(* IEC 61131-3 sources: daoli-st-library/DL_Device (part 11) *)

(* ---- FC_DL_UpsLoadRateCalc.st ---- *)
(*
 * FC_DL_UpsLoadRateCalc | C1 | DL_Device
 * 功能：UPS 负载率、N+1 冗余下的最大允许负载率与过载判定       单位：功率 [kW]、负载率 [%]、台数 [台]
 * 工况边界：模块均分假设（各模块容量相同、均流良好）；额定功率须 >0、模块数须 ≥1、冗余台数须满足 0 ≤ nRedundant < nModules；不含电池放电与效率修正
 * 代数值回代：rated=400 kW、nModules=4、nRedundant=1 → maxPct=3/4×100=75 %、允许 300 kW；load=320 kW → 320>300 → xOverload=TRUE、负载率 80 %（与 spec 回代行一致）
 * 开源溯源：clean-room 自研，未复制任何第三方代码（无外部来源）
 *)
FUNCTION FC_DL_UpsLoadRateCalc : BOOL
VAR_INPUT
    rLoadKw     : REAL := 320.0;     // 实际负载功率 | actual load power [kW]
    rRatedKw    : REAL := 400.0;     // UPS 额定功率（全模块）| UPS rated power, all modules [kW]
    nModules    : INT := 4;          // 模块总数 | total module count [台]
    nRedundant  : INT := 1;          // 冗余模块数 | redundant module count [台]
END_VAR
VAR_OUTPUT
    rLoadRatePct     : REAL;         // 负载率 | load rate [%]
    rMaxPermittedPct : REAL;         // 冗余约束下的最大允许负载率 | maximum permitted load rate under the redundancy constraint [%]
    rMaxPermittedKw  : REAL;         // 冗余约束下的最大允许负载功率 | maximum permitted load power [kW]
    xOverload        : BOOL;         // 过载（超过冗余允许值）| overload beyond the redundancy allowance
    xRedundancyOk    : BOOL;         // 冗余成立（去冗余后仍有 ≥1 台可用）| redundancy valid, at least one module remains
    xValid           : BOOL;         // 输出有效 | outputs valid
END_VAR
VAR
    xFinLoad : BOOL;                 // 负载功率有限性 | load power is finite
    xFinRated: BOOL;                 // 额定功率有限性 | rated power is finite
    nUsable  : INT;                  // 允许带载的模块数（去冗余）| usable modules after removing the redundancy [台]
    rModules : REAL;                 // 模块数实数形式 | module count as a real number [台]
END_VAR
VAR CONSTANT
    DL_ULR_PCT : REAL := 100.0;      // 百分数换算系数 | percentage factor [%]
    DL_ULR_MIN : REAL := 1.0E-9;     // 额定功率下限（防零除）| rated power lower bound [kW]
END_VAR

// 段1｜非有限闸（R19）
xFinLoad := (rLoadKw = rLoadKw) AND ((rLoadKw - rLoadKw) = 0.0);
xFinRated := (rRatedKw = rRatedKw) AND ((rRatedKw - rRatedKw) = 0.0);
IF (NOT xFinLoad) OR (NOT xFinRated) THEN
    rLoadRatePct := 0.0;             // 安全值：负载率 0 | safe value, zero load rate
    rMaxPermittedPct := 0.0;
    rMaxPermittedKw := 0.0;
    xOverload := TRUE;               // 安全值：判过载，禁止新增负载 | safe value, flagged as overload
    xRedundancyOk := FALSE;
    xValid := FALSE;
    FC_DL_UpsLoadRateCalc := FALSE;
    RETURN;
END_IF

// 段2｜域闸：额定功率入分母须 >0，模块数与冗余数须自洽
IF (rRatedKw <= DL_ULR_MIN) OR (nModules < 1) OR (nRedundant < 0) OR (nRedundant >= nModules) THEN
    rLoadRatePct := 0.0;
    rMaxPermittedPct := 0.0;
    rMaxPermittedKw := 0.0;
    xOverload := TRUE;
    xRedundancyOk := FALSE;
    xValid := FALSE;
    FC_DL_UpsLoadRateCalc := FALSE;
    RETURN;
END_IF

// 段3｜算法：maxPct = (n−nRed)/n×100；负载率 = load/rated×100
nUsable := nModules - nRedundant;
rModules := INT_TO_REAL(nModules);
rMaxPermittedPct := INT_TO_REAL(nUsable) / rModules * DL_ULR_PCT;
rMaxPermittedKw := rRatedKw * INT_TO_REAL(nUsable) / rModules;
rLoadRatePct := rLoadKw / rRatedKw * DL_ULR_PCT;

// 段4｜判定：过载与冗余度（判据同源于原始功率与台数）
xOverload := rLoadKw > rMaxPermittedKw;
xRedundancyOk := nUsable >= 1;
xValid := TRUE;
FC_DL_UpsLoadRateCalc := TRUE;
END_FUNCTION

(* ---- FC_DL_VacHoldDecayChk.st ---- *)
(*
  ============================================================
  组件名 : FC_DL_VacHoldDecayChk
  分类   : DL_Device
  功能   : 真空保持衰减校验，按保持时段内的真空度跌落求衰减率并给出泄漏报警
  复杂度 : C1
  版本   : 1.0.0
  作者   : 道莅工业代码库工厂 / R81
  日期   : 2026-11-24
  开源溯源 : clean-room（no upstream）—— 依据公开工程公式自研，未复制任何上游实现
  红线自检 : R1 无GVL/R2 无物理地址/R3 纯IEC/R4 防除零/R5 双语注释
  接口说明 :
      衰减率 = (起始真空度 - 当前真空度) / 保持时长，单位 kPa/s。
      当前真空度高于起始值属测量异常或补抽工况，衰减率按 0 处理并置 bSuspect 提示，不判泄漏。
      衰减率严格大于允许限值才置泄漏报警，等于限值视为边界可控。
  ============================================================
*)
FUNCTION FC_DL_VacHoldDecayChk : BOOL
VAR_INPUT
    bEnable     : BOOL; // 使能：TRUE 时校验 / Enable: TRUE to check
    bErr        : BOOL; // 外部故障：TRUE 时立即退出并置结果无效 / External fault: TRUE aborts with invalid result
    rVacStart_kpa : REAL; // 保持时段起始真空度 [kPa] / vacuum level at the start of the hold phase [kilopascal]
    rVacNow_kpa : REAL; // 当前实测真空度 [kPa] / current measured vacuum level [kilopascal]
    rHoldTime_s : REAL; // 保持时段已持续时长 [s] / elapsed hold phase duration [second]
    rDecayLim   : REAL; // 允许的最大衰减率 [kPa/s] / permitted maximum decay rate [kilopascal per second]
END_VAR
VAR_OUTPUT
    rDecayRate : REAL; // 实测真空衰减率，负值按 0 处理 [kPa/s] / measured vacuum decay rate, negative clamped to zero [kilopascal per second]
    rDropKpa   : REAL; // 时段内真空度跌落量 [kPa] / vacuum drop within the hold phase [kilopascal]
    bLeakAlarm : BOOL; // 泄漏报警：TRUE 表示衰减率超过限值 / leak alarm, TRUE when the decay rate exceeds the limit
    bSuspect   : BOOL; // 数据可疑：TRUE 表示当前真空度高于起始值 / suspect data, TRUE when the current vacuum is above the start value
    bValid     : BOOL; // 输出有效：TRUE 表示结果可用 / Output valid
END_VAR
VAR CONSTANT
    DL_R_MAX   : REAL := 3.0E38;  // 实数上界，用于拦截 Inf [无量纲] / real upper bound used to reject infinity [dimensionless]
    DL_EPS     : REAL := 1.0E-12; // 除零判定阈值 [无量纲] / division guard threshold [dimensionless]
    DL_ZERO    : REAL := 0.0;     // 零值常量 [无量纲] / zero constant [dimensionless]
    DL_VAC_MAX : REAL := 101.3;   // 真空度物理上限，标准大气压 [kPa] / physical upper bound of the vacuum level, standard atmosphere [kilopascal]
END_VAR
VAR
    _bFin : BOOL := FALSE; // 输入有限性判定结果 / input finiteness verdict
END_VAR

    // 段 1｜出口预置：报警位保守置 FALSE，可疑位先置 FALSE
    rDecayRate := 0.0;
    rDropKpa := 0.0;
    bLeakAlarm := FALSE;
    bSuspect := FALSE;
    bValid := FALSE;
    // 段 2｜使能闸与外部故障闸
    IF NOT bEnable THEN
        RETURN;
    END_IF;
    IF bErr THEN
        RETURN;
    END_IF;
    // 段 3｜非有限闸
    _bFin := (rVacStart_kpa = rVacStart_kpa) AND (ABS(rVacStart_kpa) <= DL_R_MAX) AND (rVacNow_kpa = rVacNow_kpa) AND (ABS(rVacNow_kpa) <= DL_R_MAX) AND (rHoldTime_s = rHoldTime_s) AND (ABS(rHoldTime_s) <= DL_R_MAX) AND (rDecayLim = rDecayLim) AND (ABS(rDecayLim) <= DL_R_MAX);
    IF NOT _bFin THEN
        RETURN;
    END_IF;
    // 段 4｜域闸：保持时长严格为正，真空度与限值不得为负
    IF (ABS(rHoldTime_s) <= DL_EPS) OR (rHoldTime_s < DL_ZERO) THEN
        RETURN;
    END_IF;
    IF (rVacStart_kpa < DL_ZERO) OR (rVacNow_kpa < DL_ZERO) OR (rDecayLim < DL_ZERO) THEN
        RETURN;
    END_IF;
    IF (rVacStart_kpa > DL_VAC_MAX) OR (rVacNow_kpa > DL_VAC_MAX) THEN
        RETURN;
    END_IF;
    // 段 5｜跌落量与衰减率
    rDropKpa := rVacStart_kpa - rVacNow_kpa;
    IF rDropKpa < DL_ZERO THEN
        bSuspect := TRUE;
        rDropKpa := DL_ZERO;
        rDecayRate := DL_ZERO;
    ELSE
        bSuspect := FALSE;
        rDecayRate := rDropKpa / rHoldTime_s;
    END_IF;
    // 段 6｜泄漏报警
    IF rDecayRate > rDecayLim THEN
        bLeakAlarm := TRUE;
    ELSE
        bLeakAlarm := FALSE;
    END_IF;
    bValid := TRUE;
    FC_DL_VacHoldDecayChk := bValid;
END_FUNCTION

(* ---- FC_DL_VacuumGenDutyCalc.st ---- *)
(*
  ============================================================
  组件名 : FC_DL_VacuumGenDutyCalc
  分类   : DL_Device
  功能   : 真空发生器占空比计算，按单周期通电时长求占空比并折算压缩空气耗量
  复杂度 : C1
  版本   : 1.0.0
  作者   : 道莅工业代码库工厂 / R81
  日期   : 2026-11-24
  开源溯源 : clean-room（no upstream）—— 依据公开工程公式自研，未复制任何上游实现
  红线自检 : R1 无GVL/R2 无物理地址/R3 纯IEC/R4 防除零/R5 双语注释
  接口说明 :
      占空比 = 通电时长 / 循环周期 * 100，限幅 0~100。
      平均耗气量 = 额定耗气量 * 占空比 / 100，单位 L/min。
      通电时长超过循环周期属参数矛盾，判无效；周期为零则无法归一，同样判无效。
  ============================================================
*)
FUNCTION FC_DL_VacuumGenDutyCalc : BOOL
VAR_INPUT
    bEnable    : BOOL; // 使能：TRUE 时计算 / Enable: TRUE to compute
    bErr       : BOOL; // 外部故障：TRUE 时立即退出并置结果无效 / External fault: TRUE aborts with invalid result
    rOnTime_s  : REAL; // 单周期内真空发生器通电时长 [s] / generator energised time within one cycle [second]
    rCycle_s   : REAL; // 循环周期总时长 [s] / total cycle duration [second]
    rAirCons   : REAL; // 通电状态下的额定耗气量 [L/min] / rated air consumption while energised [litre per minute]
END_VAR
VAR_OUTPUT
    rDutyPct   : REAL; // 真空发生器占空比，限幅 0~100 [%] / generator duty cycle clamped to 0 to 100 [percent]
    rAirUseLpm : REAL; // 折算平均耗气量 [L/min] / equivalent average air consumption [litre per minute]
    bValid     : BOOL; // 输出有效：TRUE 表示结果可用 / Output valid
END_VAR
VAR CONSTANT
    DL_R_MAX   : REAL := 3.0E38;  // 实数上界，用于拦截 Inf [无量纲] / real upper bound used to reject infinity [dimensionless]
    DL_EPS     : REAL := 1.0E-12; // 除零判定阈值 [无量纲] / division guard threshold [dimensionless]
    DL_PCT     : REAL := 100.0;   // 百分数换算系数 [无量纲] / percentage scaling factor [dimensionless]
    DL_ZERO    : REAL := 0.0;     // 零值常量 [无量纲] / zero constant [dimensionless]
    DL_TOL_S   : REAL := 0.001;   // 时长比较容差 [s] / tolerance of the duration comparison [second]
    DL_CYC_MAX : REAL := 86400.0; // 循环周期合理上限，一天 [s] / sanity upper bound of the cycle duration, one day [second]
END_VAR
VAR
    _bFin : BOOL := FALSE; // 输入有限性判定结果 / input finiteness verdict
END_VAR

    // 段 1｜出口预置
    rDutyPct := 0.0;
    rAirUseLpm := 0.0;
    bValid := FALSE;
    // 段 2｜使能闸与外部故障闸
    IF NOT bEnable THEN
        RETURN;
    END_IF;
    IF bErr THEN
        RETURN;
    END_IF;
    // 段 3｜非有限闸
    _bFin := (rOnTime_s = rOnTime_s) AND (ABS(rOnTime_s) <= DL_R_MAX) AND (rCycle_s = rCycle_s) AND (ABS(rCycle_s) <= DL_R_MAX) AND (rAirCons = rAirCons) AND (ABS(rAirCons) <= DL_R_MAX);
    IF NOT _bFin THEN
        RETURN;
    END_IF;
    // 段 4｜域闸：周期严格为正且不超过一天，通电时长与耗气量非负
    IF (ABS(rCycle_s) <= DL_EPS) OR (rCycle_s < DL_ZERO) OR (rCycle_s > DL_CYC_MAX) THEN
        RETURN;
    END_IF;
    IF (rOnTime_s < DL_ZERO) OR (rAirCons < DL_ZERO) THEN
        RETURN;
    END_IF;
    // 段 5｜通电时长不得越过周期
    IF rOnTime_s > (rCycle_s + DL_TOL_S) THEN
        RETURN;
    END_IF;
    // 段 6｜占空比与限幅
    rDutyPct := rOnTime_s / rCycle_s * DL_PCT;
    IF rDutyPct < DL_ZERO THEN
        rDutyPct := DL_ZERO;
    END_IF;
    IF rDutyPct > DL_PCT THEN
        rDutyPct := DL_PCT;
    END_IF;
    // 段 7｜平均耗气量
    rAirUseLpm := rAirCons * rDutyPct / DL_PCT;
    bValid := TRUE;
    FC_DL_VacuumGenDutyCalc := bValid;
END_FUNCTION

(* ---- FC_DL_VacuumPadForceCalc.st ---- *)
(*
  ============================================================
  组件名 : FC_DL_VacuumPadForceCalc
  分类   : DL_Device
  功能   : 真空吸盘吸附力计算，由吸盘直径与真空度求理论吸附力并按安全系数折算可用力
  复杂度 : C1
  版本   : 1.0.0
  作者   : 道莅工业代码库工厂 / R81
  日期   : 2026-11-24
  开源溯源 : clean-room（no upstream）—— 依据公开工程公式自研，未复制任何上游实现
  红线自检 : R1 无GVL/R2 无物理地址/R3 纯IEC/R4 防除零/R5 双语注释
  接口说明 :
      吸附力 F = (pi/4) * (直径/1000)^2 * (真空度*1000)，直径先由 mm 折 m，真空度由 kPa 折 Pa，结果单位 N。
      可用力 = 理论力 / 安全系数；安全系数工程常用 1.5~3，低于 1.0 视为参数错误。
      面积同时以 mm2 输出，便于与样本册的吸盘规格直接对照。
  ============================================================
*)
FUNCTION FC_DL_VacuumPadForceCalc : BOOL
VAR_INPUT
    bEnable  : BOOL; // 使能：TRUE 时计算 / Enable: TRUE to compute
    bErr     : BOOL; // 外部故障：TRUE 时立即退出并置结果无效 / External fault: TRUE aborts with invalid result
    rDia_mm  : REAL; // 吸盘有效直径 [mm] / effective pad diameter [millimetre]
    rVacKpa  : REAL; // 工作真空度 [kPa] / working vacuum level [kilopascal]
    rSafety  : REAL; // 安全系数，常用 1.5~3 [无量纲] / safety factor, typically 1.5 to 3 [dimensionless]
END_VAR
VAR_OUTPUT
    rArea_mm2 : REAL; // 吸盘有效面积 [mm2] / effective pad area [square millimetre]
    rForceN   : REAL; // 理论吸附力 [N] / theoretical holding force [newton]
    rUsableN  : REAL; // 除以安全系数后的可用吸附力 [N] / usable holding force after the safety factor [newton]
    bValid    : BOOL; // 输出有效：TRUE 表示结果可用 / Output valid
END_VAR
VAR CONSTANT
    DL_PI      : REAL := 3.14159265; // 圆周率 [无量纲] / circular constant [dimensionless]
    DL_R_MAX   : REAL := 3.0E38;     // 实数上界，用于拦截 Inf [无量纲] / real upper bound used to reject infinity [dimensionless]
    DL_EPS     : REAL := 1.0E-12;    // 除零判定阈值 [无量纲] / division guard threshold [dimensionless]
    DL_MM_TO_M : REAL := 1000.0;     // 毫米折米系数 [mm/m] / millimetre to metre factor [millimetre per metre]
    DL_KPA_TO_PA : REAL := 1000.0;   // 千帕折帕系数 [Pa/kPa] / kilopascal to pascal factor [pascal per kilopascal]
    DL_QUARTER : REAL := 0.25;       // 四分之一，用于 pi/4 折算 [无量纲] / one quarter used for the pi over four term [dimensionless]
    DL_SAFE_MIN : REAL := 1.0;       // 安全系数下界 [无量纲] / lower bound of the safety factor [dimensionless]
    DL_SAFE_MAX : REAL := 10.0;      // 安全系数上界 [无量纲] / upper bound of the safety factor [dimensionless]
    DL_VAC_MAX : REAL := 101.3;      // 真空度物理上限，标准大气压 [kPa] / physical upper bound of the vacuum level, standard atmosphere [kilopascal]
END_VAR
VAR
    _bFin  : BOOL := FALSE; // 输入有限性判定结果 / input finiteness verdict
    _rDia  : REAL := 0.0;   // 吸盘直径折算米 [m] / pad diameter in metre [metre]
    _rArea : REAL := 0.0;   // 吸盘有效面积 [m2] / effective pad area [square metre]
    _rPress : REAL := 0.0;  // 压差折算帕 [Pa] / differential pressure in pascal [pascal]
END_VAR

    // 段 1｜出口预置
    rArea_mm2 := 0.0;
    rForceN := 0.0;
    rUsableN := 0.0;
    bValid := FALSE;
    // 段 2｜使能闸与外部故障闸
    IF NOT bEnable THEN
        RETURN;
    END_IF;
    IF bErr THEN
        RETURN;
    END_IF;
    // 段 3｜非有限闸
    _bFin := (rDia_mm = rDia_mm) AND (ABS(rDia_mm) <= DL_R_MAX) AND (rVacKpa = rVacKpa) AND (ABS(rVacKpa) <= DL_R_MAX) AND (rSafety = rSafety) AND (ABS(rSafety) <= DL_R_MAX);
    IF NOT _bFin THEN
        RETURN;
    END_IF;
    // 段 4｜域闸：直径严格为正且不超过 1 m，真空度为正且不超过大气压，安全系数在合理区间
    IF (ABS(rDia_mm) <= DL_EPS) OR (rDia_mm < 0.0) OR (rDia_mm > DL_MM_TO_M) THEN
        RETURN;
    END_IF;
    IF (ABS(rVacKpa) <= DL_EPS) OR (rVacKpa < 0.0) OR (rVacKpa > DL_VAC_MAX) THEN
        RETURN;
    END_IF;
    IF (rSafety < DL_SAFE_MIN) OR (rSafety > DL_SAFE_MAX) THEN
        RETURN;
    END_IF;
    // 段 5｜面积换算
    _rDia := rDia_mm / DL_MM_TO_M;
    _rArea := DL_PI * DL_QUARTER * _rDia * _rDia;
    rArea_mm2 := DL_PI * (rDia_mm * 0.5) * (rDia_mm * 0.5);
    // 段 6｜理论吸附力：面积乘压差
    _rPress := rVacKpa * DL_KPA_TO_PA;
    rForceN := _rArea * _rPress;
    // 段 7｜安全系数除前闸后再算可用力
    IF ABS(rSafety) <= DL_EPS THEN
        RETURN;
    END_IF;
    rUsableN := rForceN / rSafety;
    bValid := TRUE;
    FC_DL_VacuumPadForceCalc := bValid;
END_FUNCTION

(* ---- FC_DL_WinderTraversePitchCalc.st ---- *)
// FC_DL_WinderTraversePitchCalc v1.0.0
// 开源溯源：clean-room 自研（族 DL_Device，ST 生态实测 0 命中，无外部代码引入）
(*
  功能: 排线节距 = 带宽·(1 − 搭接率) [mm]；换向次数 = (卷绕线速·1000/60)/(2·排线行程) [次/min]；
        排线速度 = 节距·换向次数/60 [mm/s]。此为等比近似工程式：以排线行程近似替代卷径，
        适用于定行程往复排线的稳态估算，卷径变化需上层按卷径比修正。
  邻件/码位: 与 FC_DL_FiberDiameterFromDrawRateCalc 同属拉丝后端件（卷绕面 vs 直径面）；
             16#0002_9224 = 非有限、搭接率越界或带宽/行程/线速非正拒收。
*)
FUNCTION FC_DL_WinderTraversePitchCalc : REAL
VAR_INPUT
    fStrandWidth  : REAL := 20.0;   // 丝束带宽 [mm]，域 > 0 / Strand band width [mm]
    fOverlapRatio : REAL := 0.2;    // 搭接率 [-]，域 [0, 1) / Overlap ratio
    fWinderSpeed  : REAL := 900.0;  // 卷绕线速 [m/min]，域 > 0 / Winding speed [m/min]
    fTraverseLen  : REAL := 250.0;  // 排线行程 [mm]，域 > 0 / Traverse stroke [mm]
END_VAR
VAR_OUTPUT
    fPitch          : REAL;         // 排线节距 [mm] / Traverse pitch [mm]
    fTraverseSpeed  : REAL;         // 排线速度 [mm/s] / Traverse speed [mm/s]
    fReversalPerMin : REAL;         // 每分钟换向次数 [次/min] / Reversals per minute
    bValid          : BOOL;         // 结果有效回执 [-] / Result validity receipt
    uErrorId        : UDINT;        // 事件码，0 = 无事件 / Event code
END_VAR
VAR
    fSpeedMmS    : REAL := 0.0;     // 卷绕线速 [mm/s] / Winding speed [mm/s]
    fRoundTripMm : REAL := 0.0;     // 往返行程长度 [mm] / Round-trip travel [mm]
END_VAR
// 段 0：全路径出口安全缺省 / Safe defaults on all outlets
fPitch := 0.0;                      // 节距缺省零 / Pitch default zero
fTraverseSpeed := 0.0;              // 排线速度缺省零 / Traverse speed default zero
fReversalPerMin := 0.0;             // 换向次数缺省零 / Reversal rate default zero
bValid := FALSE;                    // 有效回执预清 / Validity preset clear
uErrorId := 16#0000;                // 事件码预清 / Event code preset clear
FC_DL_WinderTraversePitchCalc := 0.0;   // 返回值缺省零（镜像节距）/ Return default zero
// 段 1：非有限闸（四入参全枚举）/ Non-finite gate over all inputs
IF (fStrandWidth <> fStrandWidth) OR (fOverlapRatio <> fOverlapRatio)
   OR (fWinderSpeed <> fWinderSpeed) OR (fTraverseLen <> fTraverseLen)
   OR (ABS(fStrandWidth) >= 3.0E38) OR (ABS(fOverlapRatio) >= 3.0E38)
   OR (ABS(fWinderSpeed) >= 3.0E38) OR (ABS(fTraverseLen) >= 3.0E38) THEN
    uErrorId := 16#0002_9224;   // 入参非有限拒收 / Non-finite input reject
    RETURN;
END_IF
// 段 2：域闸（搭接率 [0,1) 防节距非正 + 带宽/行程/线速为正，R4）/ Domain gate
IF (fOverlapRatio < 0.0) OR (fOverlapRatio >= 1.0) THEN
    uErrorId := 16#0002_9224;   // 搭接率越界，节距将非正 / Overlap ratio out of range
    RETURN;
END_IF
IF (fStrandWidth <= 1.0E-6) OR (fTraverseLen <= 1.0E-6) OR (fWinderSpeed <= 1.0E-6) THEN
    uErrorId := 16#0002_9224;   // 带宽、行程或线速非正 / Non-positive width, stroke or speed
    RETURN;
END_IF
// 段 3：主计算（节距 → 换向次数 → 排线速度）/ Main computation
fPitch := fStrandWidth * (1.0 - fOverlapRatio);                 // 节距 [mm] / Pitch
fRoundTripMm := 2.0 * fTraverseLen;                             // 往返行程 [mm] / Round-trip travel
fSpeedMmS := fWinderSpeed * 1000.0 / 60.0;                      // 卷绕线速 [mm/s] / Winding speed
fReversalPerMin := fSpeedMmS / fRoundTripMm * 60.0;             // 换向次数 [次/min] / Reversal rate
fTraverseSpeed := fPitch * fReversalPerMin / 60.0;              // 排线速度 [mm/s] / Traverse speed
// 段 4：出口闸（三输出非有限复核 + 正数复核）/ Outlet gate
IF (fPitch <> fPitch) OR (fTraverseSpeed <> fTraverseSpeed) OR (fReversalPerMin <> fReversalPerMin)
   OR (ABS(fPitch) >= 3.0E38) OR (ABS(fTraverseSpeed) >= 3.0E38) OR (ABS(fReversalPerMin) >= 3.0E38)
   OR (fPitch <= 0.0) OR (fTraverseSpeed <= 0.0) THEN
    fPitch := 0.0;              // 复核失败回缺省 / Fallback on recheck failure
    fTraverseSpeed := 0.0;      // 复核失败回缺省 / Fallback on recheck failure
    fReversalPerMin := 0.0;     // 复核失败回缺省 / Fallback on recheck failure
    uErrorId := 16#0002_9224;   // 出口复核拒收 / Output recheck reject
    RETURN;
END_IF
bValid := TRUE;                 // 有效回执 / Validity receipt
FC_DL_WinderTraversePitchCalc := fPitch;    // 返回值镜像节距 / Return mirrors pitch
END_FUNCTION

(* ---- FB_DL_AdcNoiseFloorWatch.st ---- *)
(*
  ==================================================================
  组件名 Component  : FB_DL_AdcNoiseFloorWatch
  分类   Category   : DL_Device
  前缀   Naming     : FB_DL_ ｜ b/n/u/f/t/e/st 类型前缀制（R265）
  码位   Code ID    : 16#0003_071D / 071E（故障级）｜ 16#0003_071F / 0720（信息级）
  版本   Version    : 1.0.0
  复杂度 Complexity  : 中
  功能   Purpose    : ADC 测点底噪监视：静态期窗内标准差与上限比较（接地 / 屏蔽
                      劣化、前端供电噪声的早期征兆）。
  开源溯源 Origin    : 公开公式 clean-room，参考公开测量工程口径的底噪标准差判据
                      （分类与公式借鉴，零代码复制），本件实现、闸门与码位 100% 自有。
  许可证 License    : MIT
  参考   Reference  : IEC 61131-3:2013 §6.6 算术运算符；样本标准差（n−1 分母）
                      公开统计定义
  平台   Platform   : 纯 IEC 61131-3（FOR / 四则 / SQRT / TON 无），三平台通用
  依赖   Depends    : 仅 Standard.library（SQRT 属标准内建）
  分工声明 Split     : FB_DL_SignalFrozenDetect / FB_DL_SignalStuckWatch 监视
                      不变性；FB_DL_SignalStatistics 为通用统计出口；本件为静态期
                      噪声幅度监视（动静时序由 bStatic 外部给定），四件互引（R216）。
                      SQRT 原语经派单规格授权（窗内标准差属主口径）；统计内核委托
                      不适用（流式窗口件非整段数组口径，环窗驻留数据自算）。
  归属 Ownership     : 本件无 TYPE 声明；全部引脚为 IEC 标准原生类型。
  ------------------------------------------------------------------
  边界 Boundary     :
                      一 环形窗固定容量 256（禁动态分配）；活样本恒为下标
                         0.._nFill−1（写头仅在达 _nUse 时回卷，序不变量证明同族件）；
                         标准差与均值均为序不变量，回卷不影响结果；
                      二 bStatic 变更沿全窗清零（防静 / 动混合窗污染标准差口径）；
                         nWinLen 变更沿同样清窗；
                      三 标准差两遍法（均值先行、离差平方累加在后），禁「平方和减
                         均值平方」单遍式（灾难性抵消会产生负方差或 0，SPC 经典
                         事故，写死）；除子 DINT_TO_LREAL(_nFill − 1)：_nFill < 2 →
                         不计算（判据挂起，bValid = FALSE，除零防护，R61-D4 固化）；
                      四 fNoiseLim ≤ 0 或非有限 → 组态码 071D + 三件套 + RETURN
                         结构早退（族② 判据固化，R1 教训出厂即正确）；
                      五 fMeas 非有限 → 丢弃不入窗，nNonFinite 局部计数（不外显，
                         R62-D7 口径）超窗长一半 → 故障 071E + bValid = FALSE；
                      六 判据迟滞：fNoiseStd > fNoiseLim 触发，回落
                         < fNoiseLim×(1−fHystPct/100) 复原（两方向分别定义，R146）；
                      七 bEnable = FALSE 的语义写死（FB33-4 声明行）：判据复位 +
                         fNoiseStd 冻结（纯监视件，保留读数供 HMI）；
                      八 首拍 _bInit 全量初始化；无状态机（CASE N/A，R6 标注）；
                         无定时器 / 无边沿实例（段 0 无刷新对象）；无全局、无外部
                         变量、无物理地址。
  错误码 Codes      :
    16#0003_071D【故障级】组态非法（fNoiseLim ≤ 0 / 非有限；fHystPct < 0 / 非有限）
    16#0003_071E【故障级】测量失效（非有限样本累计超过窗长一半）
    16#0003_071F【信息级】底噪超上限（bNoiseHigh = TRUE）
    16#0003_0720【信息级】窗长越域已钳位（合法 16..256）
  码位反证 Note     :
    071D 与 071E 不可合并：071D 组态即刻判（与窗内容无关），071E 需窗已建立且坏点
    累计超半窗，处置人不同（组态工程师 / 仪表工），可由 nFill 与窗状态还原（R90）；
    071F / 0720 信息级与故障级分属不同子带（R75 子带纪律），不可跨用。
  验收 Acceptance   :
    算法已证（脚本）：未跑 ｜ 编译器已证（三平台）：未跑
    V1 恒定值 → std = 0、bNoiseHigh = FALSE
    V2 注入 ±0.5 方波抖动 → std ≈ 0.5，超限触发
    V3 限值上下 5% 波动（迟滞 10%）→ 不反复跳
    V4 fNoiseLim = 0 → 组态早退；V5 _nFill = 1 → 判据挂起 bValid = FALSE
    V6 bStatic 翻转 → 清窗 nFill = 0；V7 全 NaN → 故障 071E
  修订记录 Revision  :
    2026-11-21  v1.0.0  R63 首版（批 3 · 序号 9）
  ==================================================================
*)
FUNCTION_BLOCK FB_DL_AdcNoiseFloorWatch
VAR_INPUT
    bEnable   : BOOL := TRUE;  // 使能，FALSE 时判据复位 + 标准差冻结（边界七）/ the enable, false resets the criterion and freezes the std
    fMeas     : LREAL := 0.0;  // 测点实测值 [工程单位]，必须有限 / the measured value, must be finite
    bStatic   : BOOL := FALSE; // 静态期标志（过程稳态且无操作，由调用方给）[-] / the static period flag given by the caller
    nWinLen   : DINT := 64;    // 窗长 [个]，合法域 16..256，变更沿清窗 / the window length, legal sixteen to two hundred fifty six
    fNoiseLim : LREAL := 1.0;  // 底噪上限 [工程单位]，须 > 0 / the noise ceiling, must be positive
    fHystPct  : LREAL := 10.0; // 判据迟滞 [%]，须 ≥ 0 / the criterion hysteresis in percent, non negative
END_VAR
VAR_OUTPUT
    fNoiseStd  : LREAL := 0.0;           // 窗内标准差 [工程单位] / the window standard deviation
    bNoiseHigh : BOOL := FALSE;          // 底噪超限判据（带迟滞）[-] / the noise high criterion with hysteresis
    nFill      : DINT := 0;              // 窗填充数 [个] / the filled count
    bValid     : BOOL := FALSE;          // 判据可用 [-] / the criterion is usable
    eErr       : UDINT := 16#0000_0000;  // 错误码，0 = 正常 / the error code, zero is ok
    bError     : BOOL := FALSE;          // 故障标志（故障级码同拍置位，R45 配对）/ the fault flag raised with a fault level code
END_VAR
VAR
    _bInit     : BOOL := FALSE;              // 首拍初始化标志（R310 / FB50-2）/ the first scan flag
    _afWin     : ARRAY[0..255] OF LREAL;     // 采样环形窗 [工程单位]，固定容量 256 / the fixed capacity ring of samples
    _nHead     : DINT := 0;                  // 环形窗写头 [下标] / the ring write head
    _nFill     : DINT := 0;                  // 环形窗填充计数 [个] / the ring filled count
    _nUse      : DINT := 64;                 // 钳位后的窗长 [个] / the clamped window length
    _nUsePrev  : DINT := 0;                  // 上拍窗长快照 [个]，置 0 使首拍必触发清窗 / the previous length
    _bStaticPrev : BOOL := FALSE;            // 上拍静态期快照 [-] / the previous static flag
    _nClrIdx   : DINT := 0;                  // 清窗遍历索引 [下标] / the clearing traversal index
    _nSumIdx   : DINT := 0;                  // 统计遍历索引 [下标] / the statistics traversal index
    _nNonFinite: DINT := 0;                  // 非有限丢弃计数 [个]（仅局部留档，不外显，R62-D7 口径）/ the dropped non finite count, local only and never exposed
    _fSum      : LREAL := 0.0;               // 窗内样本和 [工程单位] / the window sample sum
    _fMean     : LREAL := 0.0;               // 窗内均值（两遍法第一遍）[工程单位] / the window mean of the first pass
    _fSqSum    : LREAL := 0.0;               // 离差平方和（两遍法第二遍）[工程单位²] / the squared deviation sum of the second pass
    _fStdUse   : LREAL := 0.0;               // 标准差工作副本 [工程单位] / the working standard deviation
    _fVar      : LREAL := 0.0;               // 样本方差（n−1 分母）[工程单位²] / the sample variance
    _bNoiseL   : BOOL := FALSE;              // 底噪超限迟滞状态（跨拍保持）/ the noise high hysteresis state
    _bCfgBad   : BOOL := FALSE;              // 组态非法标记（逐拍重算）/ the configuration fault flag
    _bWinClamp : BOOL := FALSE;              // 窗长钳位标记（逐拍重算，信息级 0720）/ the window clamp flag
    _bMeasBad  : BOOL := FALSE;              // 测量失效标记（逐拍重算）/ the measurement failure flag
    _bFinLim   : BOOL := FALSE;              // 上限有限闸结果（逐拍重算）/ the limit finiteness gate result
    _bFinHyst  : BOOL := FALSE;              // 迟滞有限闸结果（逐拍重算）/ the hysteresis finiteness gate result
    _bFinMeas  : BOOL := FALSE;              // 样本有限闸结果（逐拍重算）/ the sample finiteness gate result
END_VAR  // R64 结构补齐：VAR 段缺失的 END_VAR（门禁机械修复）
VAR CONSTANT
    DL_ANF_WMAX  : DINT := 256;      // 窗容量上界 [个]，与数组容量一致 / the capacity aligned with the array
    DL_ANF_WMIN  : DINT := 16;       // 窗长下界 [个] / the window floor
    DL_ANF_ZERO  : LREAL := 0.0;     // 实数零常量 [工程单位] / the real zero constant
    DL_ANF_PCT   : LREAL := 100.0;  // 百分比换算系数 [%] / the percentage scaling factor
    DL_ANF_ONE   : DINT := 1;        // 整型一常量 [个] / the integer one constant
    DL_ANF_TWO   : DINT := 2;        // 整型二常量 [个]（方差最少样本）/ the integer two constant, the minimum for a variance
    DL_ANF_ZEROI : DINT := 0;        // 整型零常量 [个] / the integer zero constant
    DL_ANF_HALF  : LREAL := 2.0;     // 半窗判据除子 [−] / the half window criterion divisor
END_VAR

// 段 0｜本件无定时器与边沿实例（纯统计监视器，R6 标注 N/A），无刷新对象 / segment 0, no timers and no edge instances exist here

// 段 1｜首拍初始化（FB50-2）/ segment 1, the first scan init
IF NOT _bInit THEN // 首拍一拍 / the first scan
    _bInit := TRUE; // 置首拍标志 / raise the first scan flag
    _nFill := DL_ANF_ZEROI; // 填充计数显式清零 / clear the filled count explicitly
    _nHead := DL_ANF_ZEROI; // 写头显式清零 / clear the write head explicitly
    _fSum := DL_ANF_ZERO; // 窗和显式清零 / clear the sum explicitly
    _nUsePrev := DL_ANF_ZEROI; // 窗长快照置 0，使段 3 变更沿必然触发一次清窗 / zero the snapshot so the change edge clears once
    _bStaticPrev := bStatic; // 静态期快照对齐首拍值（防首拍误清窗）/ align the static snapshot to avoid a spurious clear
    _bNoiseL := FALSE; // 迟滞状态显式清零 / clear the hysteresis state explicitly
    _nNonFinite := DL_ANF_ZEROI; // 非有限计数显式清零 / clear the non finite count explicitly
    FOR _nClrIdx := DL_ANF_ZEROI TO DL_ANF_WMAX - DL_ANF_ONE DO // 有界遍历全容量 / the bounded traversal over the full capacity
        _afWin[_nClrIdx] := DL_ANF_ZERO; // 窗元素逐项清零 / zero every window element
    END_FOR
END_IF

// 段 2｜组态域闸（边界四，族② 判据：全部限值逐个点名，R272）/ segment 2, the configuration gates
_bFinLim := (fNoiseLim = fNoiseLim) AND ((fNoiseLim - fNoiseLim) = (fNoiseLim - fNoiseLim)); // 上限有限 / the ceiling is finite
_bFinHyst := (fHystPct = fHystPct) AND ((fHystPct - fHystPct) = (fHystPct - fHystPct)); // 迟滞有限 / the hysteresis is finite
_bCfgBad := (NOT _bFinLim) OR (fNoiseLim <= DL_ANF_ZERO) OR (NOT _bFinHyst) OR (fHystPct < DL_ANF_ZERO); // 组态非法 / an illegal configuration
IF _bCfgBad THEN // 组态非法：结构早退（出口三件套 + RETURN，除法段不可达）/ an illegal configuration exits structurally
    fNoiseStd := _fStdUse; // 标准差取最近有效值 [工程单位]（禁自赋值出口，R261）/ the std takes the last valid value instead of a self assignment
    bNoiseHigh := FALSE; // 判据复位 / the criterion resets
    nFill := _nFill; // 填充计数照实出口 [个] / the fill count as is
    bValid := FALSE; // 判据不可用 / the criterion is not usable
    eErr := 16#0003_071D; // 故障级：组态非法 / fault grade, an illegal configuration
    bError := TRUE; // 同拍置故障标志（R45 配对）/ raise the fault flag on the same scan
    RETURN; // 结构早退 / the structural early exit
END_IF

// 段 3｜窗长钳位与变更沿 / 静态期变更沿全窗清零（边界二）/ segment 3, the window clamp and the change edge clears
_bWinClamp := FALSE; // 钳位标记预清零（单拍信息位，段 8 映射）/ preset the clamp flag false
_bMeasBad := FALSE; // 测量失效标记预清零 / preset the failure flag false
_nUse := nWinLen; // 窗长接管 [个] / take the window length
IF (_nUse < DL_ANF_WMIN) OR (_nUse > DL_ANF_WMAX) THEN // 窗长越域 / the length is out of the domain
    _bWinClamp := TRUE; // 置钳位标记（信息级 0720）/ raise the clamp flag
    IF _nUse < DL_ANF_WMIN THEN // 下界钳位 / the floor clamp
        _nUse := DL_ANF_WMIN; // 钳到下界 [个] / clamp to the floor
    ELSE // 上界钳位 / the ceiling clamp
        _nUse := DL_ANF_WMAX; // 钳到容量 [个] / clamp to the capacity
    END_IF
END_IF
IF (_nUse <> _nUsePrev) OR (bStatic <> _bStaticPrev) THEN // 窗长或静态期变更沿（含首拍）/ the length or the static flag changed
    _nHead := DL_ANF_ZEROI; // 写头回零 / reset the write head
    _nFill := DL_ANF_ZEROI; // 填充计数回零 / reset the filled count
    _fSum := DL_ANF_ZERO; // 窗和回零 / reset the sum
    _nNonFinite := DL_ANF_ZEROI; // 非有限计数回零 / reset the non finite count
    FOR _nClrIdx := DL_ANF_ZEROI TO DL_ANF_WMAX - DL_ANF_ONE DO // 有界遍历全容量 / the bounded traversal over the full capacity
        _afWin[_nClrIdx] := DL_ANF_ZERO; // 窗元素逐项清零（禁静动混合窗） / zero every element so no mixed window remains
    END_FOR
    _nUsePrev := _nUse; // 快照本拍窗长 / snapshot the length
    _bStaticPrev := bStatic; // 快照本拍静态期 / snapshot the static flag
END_IF

// 段 4｜失能分支：判据复位 + 标准差冻结（边界七声明行）/ segment 4, the disabled branch
IF NOT bEnable THEN // 失能 / disabled
    fNoiseStd := _fStdUse; // 标准差冻结最近有效值 [工程单位] / freeze the last valid std
    bNoiseHigh := FALSE; // 判据复位 / the criterion resets
    nFill := _nFill; // 填充计数照实出口 [个] / the fill count as is
    bValid := FALSE; // 失能即不可用 / the criterion is not usable while disabled
    bError := FALSE; // 失能不是故障 / a disabled device is not a fault
    eErr := 16#0000_0000; // 失能不发码 / no code is emitted while disabled
    RETURN; // 早退，窗保留 / early return with the window kept
END_IF

// 段 5｜样本入窗（非有限丢弃并计数，边界五）/ segment 5, push the sample or count the drop
_bFinMeas := (fMeas = fMeas) AND ((fMeas - fMeas) = (fMeas - fMeas)); // 样本有限 / the sample is finite
IF bStatic AND _bFinMeas THEN // 静态期且样本有限才入窗（动态期样本不进底噪窗）/ only a finite sample of a static period enters the noise window
    _fSum := _fSum - _afWin[_nHead] + fMeas; // 滑窗和更新 [工程单位] / update the sliding sum
    _afWin[_nHead] := fMeas; // 本拍样本入环 [工程单位] / push the sample
    _nHead := _nHead + DL_ANF_ONE; // 写头推进 / advance the head
    IF _nHead >= _nUse THEN // 回卷（按钳位窗长）/ wrap by the clamped length
        _nHead := DL_ANF_ZEROI; // 写头回零 / reset the head
    END_IF
    IF _nFill < _nUse THEN // 窗未满才累加 / count only while not full
        _nFill := _nFill + DL_ANF_ONE; // 填充计数推进 [个] / advance the filled count
    END_IF
ELSIF bStatic THEN // 静态期但样本非有限：丢弃计数 / a static period sample is broken, dropped and counted
    _nNonFinite := _nNonFinite + DL_ANF_ONE; // 非有限计数推进 [个] / advance the non finite count
END_IF
IF DINT_TO_LREAL(_nNonFinite) > (DINT_TO_LREAL(_nUse) / DL_ANF_HALF) THEN // 非有限累计超窗长一半（边界五）/ the non finite count exceeds half the window
    _bMeasBad := TRUE; // 置测量失效标记（码 071E）/ raise the failure flag
END_IF
nFill := _nFill; // 填充计数出口 [个] / the fill count outlet

// 段 6｜均值与标准差两遍法（边界三：除子 _nFill−1，_nFill < 2 判据挂起）/ segment 6, the two pass mean and standard deviation
IF _nFill >= DL_ANF_TWO THEN // 除子已证 ≥ 1（禁裸除子）/ the divisor is proven at least one
    _fMean := _fSum / DINT_TO_LREAL(_nFill); // 第一遍：窗均值 [工程单位] / the first pass mean
    _fSqSum := DL_ANF_ZERO; // 离差平方和清零 [工程单位²] / clear the squared deviation sum
    FOR _nSumIdx := DL_ANF_ZEROI TO _nFill - DL_ANF_ONE DO // 有界遍历活样本（上界已证 ≤ 256）/ the bounded traversal over the live samples
        _fSqSum := _fSqSum + ((_afWin[_nSumIdx] - _fMean) * (_afWin[_nSumIdx] - _fMean)); // 第二遍：离差平方累加 [工程单位²] / the second pass accumulates the squared deviations
    END_FOR
    _fVar := _fSqSum / DINT_TO_LREAL(_nFill - DL_ANF_ONE); // 样本方差（n−1 分母）[工程单位²] / the sample variance with the n minus one divisor
    IF _fVar < DL_ANF_ZERO THEN // 负方差兜底（两遍法下理论上不可达，防御保留）/ a negative variance, unreachable by theory, kept as a defence
        _fVar := DL_ANF_ZERO; // 方差钳零 [工程单位²] / clamp the variance to zero
    END_IF
    _fStdUse := SQRT(_fVar); // 标准差 [工程单位]，SQRT 属主口径见分工声明 / the standard deviation
ELSE // 样本不足：判据挂起 / too few samples, the criterion suspends
    fNoiseStd := _fStdUse; // 标准差保持最近有效值 [工程单位] / keep the last valid std
    bNoiseHigh := FALSE; // 判据复位 / the criterion resets
    bValid := FALSE; // 判据不可用（_nFill < 2，边界三）/ the criterion is not usable
    eErr := 16#0000_0000; // 挂起不是故障 / a suspension is not a fault
    bError := FALSE; // 无故障 / no fault
    RETURN; // 早退，禁除零 / early return, no division is reached
END_IF

// 段 7｜底噪判据迟滞（边界六，两方向分别定义，R146）/ segment 7, the noise criterion hysteresis
IF NOT _bNoiseL THEN // 未报警态 / the released state
    IF _fStdUse > fNoiseLim THEN // 超过上限 / above the ceiling
        _bNoiseL := TRUE; // 置迟滞状态 / set the hysteresis state
    END_IF
ELSE // 已报警态 / the tripped state
    IF _fStdUse < (fNoiseLim * (DL_ANF_PCT - fHystPct) / DL_ANF_PCT) THEN // 回落低于上限减迟滞 / below the ceiling minus the hysteresis
        _bNoiseL := FALSE; // 复原 / release
    END_IF
END_IF

// 段 8｜统一出口（单拍位映射 + 信息级重算，R187 / FB51-8）/ segment 8, the unified outlet
fNoiseStd := _fStdUse; // 标准差出口 [工程单位] / the std outlet
bNoiseHigh := _bNoiseL; // 判据出口（迟滞状态派生）/ the criterion outlet
bValid := (NOT _bMeasBad); // 判据可用（无测量失效）/ usable without a measurement failure
IF _bMeasBad THEN // 测量失效（故障级优先）/ the measurement failed
    bValid := FALSE; // 判据不可用 / the criterion is not usable
    bError := TRUE; // 故障位置位 / raise the fault bit
    eErr := 16#0003_071E; // 故障级：测量失效 / fault grade, the measurement failed
ELSIF _bNoiseL THEN // 底噪超限（信息级）/ the noise is high, informational
    bError := FALSE; // 信息级不置故障位 / the informational code never raises the fault bit
    eErr := 16#0003_071F; // 信息级：底噪超上限 / informational, the noise is over the ceiling
ELSIF _bWinClamp THEN // 窗长钳位（信息级）/ the length clamp, informational
    bError := FALSE; // 信息级不置故障位 / no fault bit
    eErr := 16#0003_0720; // 信息级：窗长越域已钳位 / informational, the length was clamped
ELSE // 无事件 / no event
    bError := FALSE; // 无故障 / no fault
    eErr := 16#0000_0000; // 正常 / ok
END_IF
END_FUNCTION_BLOCK

(* ---- FB_DL_AhuFilterDpBank.st ---- *)
// =====================================================================
// FB_DL_AhuFilterDpBank.st
// 空调箱 4 段过滤器压差四级分档（迟滞 + 各段独立去抖 + 低风量冻结）
// AHU 4-stage filter dP grading with per-stage debounce and hysteresis
// 所属子库: DL_Device    版本: v1.0.0    兼容: CODESYS V3.5+ / TwinCAT 3 / 汇川 InoProShop
// 码位: 16#0003_03D9 ~ 16#0003_03DD (本件独占 5 槽, 勿复用)
// 溯源: 道莅 clean-room 防御性实现
//       来源组标签: hvac, filter-monitoring, dp-grading, hysteresis, debounce
// 枚举属主: E_DL_FilterStage —— 本文件为全库唯一属主, 其他件只引用不重声明
// 修改记录: R30 初版 (ROUND_PLAN_R30 序 1, 由 R29 隔离底稿返修入册)
//           返修要点: 共享单实例去抖定时器改为 4 温区独立实例数组 aTonDeb,
//           每扫描周期无条件刷新全部 4 个 TON 实例, 候选作废显式复位;
//           任一区间切换去抖期间其他区间计时不被复位/冻结(验收点);
//           码位由作废段 03C5~03C9 重排为实测游标新段 03D9~03DD
// =====================================================================
// ---------------------------------------------------------------------
// 枚举定义: E_DL_FilterStage (全库唯一属主, 其他件只引用不重声明)
// ---------------------------------------------------------------------
TYPE E_DL_FilterStage :
(
    eClean,         // 洁净档 / Clean stage
    eEarly,         // 初堵档 / Early clog stage
    eMid,           // 中堵档 / Mid clog stage
    eChange,        // 更换档 / Change stage
    eSensorFault    // 传感器故障档 / Sensor fault stage
);
END_TYPE

FUNCTION_BLOCK FB_DL_AhuFilterDpBank
VAR_INPUT
    bEnable        : BOOL  := FALSE;   // 使能 / Enable
    afDp_Pa        : ARRAY[1..4] OF REAL;   // 各段压差 0~2000 Pa / Stage dP [Pa]
    afDpEarly_Pa   : ARRAY[1..4] OF REAL;   // 各段初堵阈值 10~500 Pa / Early clog threshold [Pa]
    afDpChange_Pa  : ARRAY[1..4] OF REAL;   // 各段更换阈值 20~1000 Pa / Change threshold [Pa]
    fHyst_Pa       : REAL  := 10.0;    // 迟滞回差 0~100 Pa / Hysteresis band [Pa]
    fDpMax_Pa      : REAL  := 1500.0;  // 传感器量程上限 >0 Pa / Sensor range limit [Pa]
    fFanPct        : REAL  := 0.0;     // 风机输出 0~100 百分比 / Fan duty [pct]
    fFanMinPct     : REAL  := 20.0;    // 判定最低风量 0~100 百分比 / Min fan duty for judging [pct]
    tDebounce      : TIME  := T#5S;    // 去抖时长 T#100MS~T#120S / Debounce duration [s]
END_VAR
VAR_OUTPUT
    aeStage        : ARRAY[1..4] OF E_DL_FilterStage;  // 各段档位 / Stage level per section
    auMaxStage     : USINT := 0;       // 全箱最高档 0~3 / Max stage of bank 0..3
    bChangeReq     : BOOL := FALSE;    // 更换请求 / Filter change required
    bFrozen        : BOOL := FALSE;    // 低风量冻结标志 / Frozen by low airflow
    eErr           : UDINT := 16#0003_03D9;  // 错误码 / Error code
END_VAR
VAR
    aTonDeb        : ARRAY[1..4] OF TON;   // 各段独立去抖定时器, 每拍无条件刷新 / Per-stage debounce timers, refreshed every cycle
    aPendStage     : ARRAY[1..4] OF E_DL_FilterStage;  // 各段候选档位 / Pending stage per section
    aPendActive    : ARRAY[1..4] OF BOOL;  // 各段候选有效标记 / Pending active flag per section
    eAbtCode       : UDINT := 16#0003_03D9;  // 本拍守卫闸中止码 / Abort code of this cycle
    bAbort         : BOOL := FALSE;    // 守卫闸中止标记 / Gate abort flag
    bSensorFlt     : BOOL := FALSE;    // 任一段传感器故障标记 / Any-stage sensor fault flag
    uZi            : INT   := 1;       // 1..4 数组下标 / Array subscript 1..4
    eTarget        : E_DL_FilterStage := E_DL_FilterStage.eClean;  // 本拍目标档 / Target stage this cycle
    uMaxTmp        : USINT := 0;       // 最高档临时量 / Max stage temporary
    tDebS          : REAL  := 0.0;     // 去抖秒值 / Debounce seconds [s]
    xFirstScan     : BOOL  := TRUE;    // 首扫标记 / First-scan flag
END_VAR

// ---------------------------------------------------------------------
// 代码位表（本件独占, 勿复用）:
//   16#0003_03D9 信息 分档正常
//   16#0003_03DA 故障 去抖时长非法或任一标量/数组输入非有限（本拍冻结保持, 非锁存, 恢复合法输入即解除）
//   16#0003_03DB 故障 阈值组态非法（量程上限不大于 0 或任一段初堵阈值不低于更换阈值）
//   16#0003_03DC 信息 低风量冻结（风机输出低于判定下限, 档位保持不推进）
//   16#0003_03DD 故障 任一段压差超量程或为负, 该段落传感器故障档
// ---------------------------------------------------------------------

// ---- 去抖秒值换算 / Debounce seconds conversion ----
tDebS := TIME_TO_REAL(tDebounce) / 1000.0;  // 毫秒换算秒 / Convert ms to seconds [s]

// ---- 守卫闸 1: 标量输入非有限与去抖时长合法域 / Gate 1: scalar finite and debounce range ----
bAbort    := FALSE;                 // 中止标记复位 / Reset abort flag
eAbtCode  := 16#0003_03D9;          // 中止码复位 / Reset abort code
IF (tDebounce = T#0MS) OR (tDebS < 0.1) OR (tDebS > 120.0)
   OR (fHyst_Pa <> fHyst_Pa) OR (ABS(fHyst_Pa) >= 1.0E12)
   OR (fDpMax_Pa <> fDpMax_Pa) OR (ABS(fDpMax_Pa) >= 1.0E12)
   OR (fFanPct <> fFanPct) OR (ABS(fFanPct) >= 1.0E12)
   OR (fFanMinPct <> fFanMinPct) OR (ABS(fFanMinPct) >= 1.0E12) THEN
    bAbort  := TRUE;                // 置中止 / Set abort
    eAbtCode := 16#0003_03DA;       // 码 03DA / Code 03DA
END_IF

// ---- 守卫闸 2: 逐段压差与阈值非有限判界 / Gate 2: per-stage finite check ----
IF NOT bAbort THEN
    FOR uZi := 1 TO 4 DO
        IF (afDp_Pa[uZi] <> afDp_Pa[uZi]) OR (ABS(afDp_Pa[uZi]) >= 1.0E12)
           OR (afDpEarly_Pa[uZi] <> afDpEarly_Pa[uZi]) OR (ABS(afDpEarly_Pa[uZi]) >= 1.0E12)
           OR (afDpChange_Pa[uZi] <> afDpChange_Pa[uZi]) OR (ABS(afDpChange_Pa[uZi]) >= 1.0E12) THEN
            bAbort   := TRUE;           // 置中止 / Set abort
            eAbtCode := 16#0003_03DA;   // 码 03DA / Code 03DA
        END_IF
    END_FOR
END_IF

// ---- 守卫闸 3: 阈值组态合法性 / Gate 3: threshold configuration ----
IF NOT bAbort THEN
    IF fDpMax_Pa <= 0.0 THEN
        bAbort   := TRUE;           // 量程非法 / Illegal range
        eAbtCode := 16#0003_03DB;   // 码 03DB / Code 03DB
    END_IF
END_IF
IF NOT bAbort THEN
    FOR uZi := 1 TO 4 DO
        IF afDpEarly_Pa[uZi] >= afDpChange_Pa[uZi] THEN
            bAbort   := TRUE;           // 阈值倒置 / Inverted thresholds
            eAbtCode := 16#0003_03DB;   // 码 03DB / Code 03DB
        END_IF
    END_FOR
END_IF

// ---- 首扫初始化 / First-scan initialization ----
IF xFirstScan THEN
    FOR uZi := 1 TO 4 DO
        aeStage[uZi]     := E_DL_FilterStage.eClean;    // 初始洁净档 / Init clean stage
        aPendStage[uZi]  := E_DL_FilterStage.eClean;    // 候选初始 / Pending init
        aPendActive[uZi] := FALSE;  // 候选无效 / Pending inactive
    END_FOR
    xFirstScan := FALSE;        // 清首扫标记 / Clear first-scan flag
END_IF

// ---- 低风量冻结与中止冻结推导 / Low-airflow freeze and abort freeze ----
IF bAbort THEN
    bFrozen := TRUE;            // 守卫闸中止按安全冻结处理 / Abort treated as safe freeze
ELSIF fFanPct < fFanMinPct THEN
    bFrozen := TRUE;            // 低风量冻结 / Low airflow freeze
ELSE
    bFrozen := FALSE;           // 正常非冻结 / Normal not frozen
END_IF

// ---- 逐段目标档计算与候选登记（不在此处调定时器）/ Per-stage target and pending registration ----
IF NOT bAbort AND NOT bFrozen THEN
    bSensorFlt := FALSE;        // 传感器故障标记复位 / Reset sensor fault flag
    bChangeReq := FALSE;        // 更换请求复位 / Reset change request
    FOR uZi := 1 TO 4 DO
        // 传感器故障判: 超量程或负压差 / Sensor fault: over-range or negative dP
        IF (afDp_Pa[uZi] > fDpMax_Pa) OR (afDp_Pa[uZi] < 0.0) THEN
            aeStage[uZi]     := E_DL_FilterStage.eSensorFault;  // 落传感器故障档 / Sensor fault stage
            aPendActive[uZi] := FALSE;  // 候选作废 / Pending void
            bSensorFlt := TRUE;         // 置传感器故障 / Set sensor fault
            bChangeReq := TRUE;         // 故障档也需现场处置 / Fault stage requests action
        ELSE
            // 双阈值迟滞分档: 严格大于阈值才切档, 恰好等于阈值保持原档 / Strict-greater hysteresis grading
            CASE aeStage[uZi] OF
                E_DL_FilterStage.eClean:        // 当前洁净 / Currently clean
                    IF afDp_Pa[uZi] > (afDpEarly_Pa[uZi] + fHyst_Pa) THEN
                        eTarget := E_DL_FilterStage.eEarly;     // 越升档阈值 → 初堵 / Above rise threshold
                    ELSE
                        eTarget := E_DL_FilterStage.eClean;     // 保持 / Hold
                    END_IF
                E_DL_FilterStage.eEarly:        // 当前初堵 / Currently early
                    IF afDp_Pa[uZi] > (afDpChange_Pa[uZi] + fHyst_Pa) THEN
                        eTarget := E_DL_FilterStage.eChange;    // 越更换阈值 / Above change threshold
                    ELSIF afDp_Pa[uZi] < (afDpEarly_Pa[uZi] - fHyst_Pa) THEN
                        eTarget := E_DL_FilterStage.eClean;     // 回落洁净 / Fall back clean
                    ELSE
                        eTarget := E_DL_FilterStage.eEarly;     // 保持 / Hold
                    END_IF
                E_DL_FilterStage.eMid:          // 当前中堵 / Currently mid
                    IF afDp_Pa[uZi] > (afDpChange_Pa[uZi] + fHyst_Pa) THEN
                        eTarget := E_DL_FilterStage.eChange;    // 越更换阈值 / Above change threshold
                    ELSIF afDp_Pa[uZi] < (afDpEarly_Pa[uZi] - fHyst_Pa) THEN
                        eTarget := E_DL_FilterStage.eClean;     // 回落洁净 / Fall back clean
                    ELSE
                        eTarget := E_DL_FilterStage.eMid;       // 保持 / Hold
                    END_IF
                E_DL_FilterStage.eChange:       // 当前更换档 / Currently change
                    IF afDp_Pa[uZi] < (afDpChange_Pa[uZi] - fHyst_Pa) THEN
                        eTarget := E_DL_FilterStage.eMid;       // 回落中堵 / Fall back mid
                    ELSE
                        eTarget := E_DL_FilterStage.eChange;    // 保持 / Hold
                    END_IF
                E_DL_FilterStage.eSensorFault:  // 故障档: 压差恢复量程内后按洁净档重新进入 / Fault holds, re-enter via grading
                    eTarget := E_DL_FilterStage.eClean;     // 目标回洁净档, 去抖后切换 / Target clean, switch after debounce
                ELSE                            // 非法档位拦截 / Illegal stage interception
                    eTarget := E_DL_FilterStage.eSensorFault;   // 落故障档 / Fall to fault stage
            END_CASE

            // 候选登记: 目标与当前不同才登记 / Register pending only if target differs
            IF eTarget <> aeStage[uZi] THEN
                IF (NOT aPendActive[uZi]) OR (aPendStage[uZi] <> eTarget) THEN
                    aPendStage[uZi]  := eTarget;    // 登记新候选 / Register new candidate
                    aPendActive[uZi] := TRUE;       // 候选有效 / Pending active
                END_IF
            ELSE
                aPendActive[uZi] := FALSE;      // 目标即当前档, 候选作废 / Target equals current, void
            END_IF
        END_IF

        // 更换档请求判 / Change stage request check
        IF aeStage[uZi] = E_DL_FilterStage.eChange THEN
            bChangeReq := TRUE;     // 任一段处于更换档 / Any stage at change
        END_IF
    END_FOR
ELSE
    bSensorFlt := FALSE;            // 冻结/中止拍不重推传感器判据 / No sensor re-judge on frozen cycle
    bChangeReq := FALSE;            // 冻结拍不置更换请求 / No change request on frozen cycle
END_IF

// ---- 4 个去抖定时器无条件周期刷新（本 FOR 循环每拍必执行全部 4 个实例,
//      不放进任何 IF 分支; 候选作废分支传 IN 为假显式复位而不是跳过调用）
//      Unconditional refresh of all 4 TON instances every cycle ----
FOR uZi := 1 TO 4 DO
    IF (NOT bAbort) AND (NOT bFrozen) AND aPendActive[uZi] AND (aPendStage[uZi] <> aeStage[uZi]) THEN
        aTonDeb[uZi](IN := TRUE, PT := tDebounce);  // 本拍继续计时 / Keep timing this cycle
        IF aTonDeb[uZi].Q THEN
            aeStage[uZi] := aPendStage[uZi];        // 去抖通过, 档位切换 / Switch after debounce
            aPendActive[uZi] := FALSE;              // 候选完成 / Pending done
        END_IF
    ELSE
        aPendActive[uZi] := FALSE;                  // 候选作废 / Pending void
        aTonDeb[uZi](IN := FALSE, PT := tDebounce); // 候选作废显式复位 / Explicit reset on void
    END_IF
END_FOR

// ---- 最高档统计（只统计非传感器故障段）/ Max stage excluding sensor-fault sections ----
uMaxTmp := 0;                   // 临时量复位 / Reset temporary
FOR uZi := 1 TO 4 DO
    IF aeStage[uZi] <> E_DL_FilterStage.eSensorFault THEN
        CASE aeStage[uZi] OF
            E_DL_FilterStage.eClean:    // 档 0 / Stage 0
                uMaxTmp := uMaxTmp;     // 保持 0 / Keep 0
            E_DL_FilterStage.eEarly:    // 档 1 / Stage 1
                IF uMaxTmp < 1 THEN
                    uMaxTmp := 1;       // 升到 1 / Raise to 1
                END_IF
            E_DL_FilterStage.eMid:      // 档 2 / Stage 2
                IF uMaxTmp < 2 THEN
                    uMaxTmp := 2;       // 升到 2 / Raise to 2
                END_IF
            E_DL_FilterStage.eChange:   // 档 3 / Stage 3
                uMaxTmp := 3;           // 升到 3 / Raise to 3
            ELSE                        // 兜底: 非法档不计入 / Fallback: illegal stage not counted
                uMaxTmp := uMaxTmp;     // 保持 / Keep
        END_CASE
    END_IF
END_FOR
auMaxStage := uMaxTmp;          // 输出最高档 / Output max stage

// ---- 错误码仲裁（每拍重算, 非锁存, 恢复合法输入即解除）/ Error arbitration recomputed each cycle ----
IF bAbort THEN
    eErr := eAbtCode;           // 守卫闸中止码优先 / Gate abort code first
ELSIF bSensorFlt THEN
    eErr := 16#0003_03DD;       // 传感器故障 / Sensor fault
ELSIF bFrozen THEN
    eErr := 16#0003_03DC;       // 低风量冻结 / Low airflow freeze
ELSE
    eErr := 16#0003_03D9;       // 分档正常 / Grading normal
END_IF

END_FUNCTION_BLOCK

(* ---- FB_DL_AirCompressorLoadUnload.st ---- *)
(*
  Name        : FB_DL_AirCompressorLoadUnload
  Category    : DL_Device
  Version     : 1.0.0
  Purpose     : 空压机加卸载调压：压力带双阈迟滞加卸载切换，加载最小驻留防短周期振荡，卸载超时置维护级告警不自动停机；/ Air compressor load/unload pressure control: dual-threshold hysteresis switching, minimum load dwell against short cycling, unload timeout raising a maintenance-level warning without auto stop
  溯源        : 借 lbp-basic-process 与行业池的调压组织，clean-room 实现
  Boundary    : ① 压力带组态闸：加载阈 < 卸载阈否则锁存故障（相等不立）；
                ② 双阈迟滞直比（加载阈/卸载阈比较，禁浮点等值）；
                ③ 卸载持续 > 卸载超时 → 置维护级告警（bMaintWarn 锁存至复位沿，不自动停机不迁故障相，属主边界）；
                ④ 加载最小驻留防短周期振荡：驻留期内卸载请求暂存不丢（驻留满即执行）；
                ⑤ 压力传感器非有限 → 保持当前负载态 + bSensorBad 当拍出口（不切态防误动作）；
                ⑥ 本件为命令层，不直接驱动接触器（属主边界，出加/卸载命令信号）。
*)
TYPE E_DL_AclState :
(
    eIdle   := 0,                            (* 未使能（命令全停） / Idle, commands off *)
    eLoad   := 10,                           (* 加载相 / Loading *)
    eUnload := 20,                           (* 卸载相 / Unloading *)
    eFault  := 90                            (* 故障锁存相 / Fault latched *)
);
END_TYPE

TYPE E_DL_AclCause :
(
    eNone      := 0,                         (* 无成因 / No cause *)
    eCfgIllegal:= 1,                        (* 组态非法：压力带阈值倒挂 / Illegal config *)
    eUnloadTime:= 2,                        (* 维护级：卸载超时（不置 bError，边界③） / Maintenance: unload timeout *)
    ePhaseBad  := 3                         (* 非法相位兜底 / Illegal phase fallback *)
);
END_TYPE

FUNCTION_BLOCK FB_DL_AirCompressorLoadUnload
VAR_INPUT
    fPress   : REAL := 0.0;                  (* 储气罐压力 [bar] / Receiver pressure *)
    fLoadTh  : REAL := 6.0;                  (* 加载阈（下限），域 < 卸载阈 [bar] / Load threshold *)
    fUnloadTh: REAL := 8.0;                  (* 卸载阈（上限）[bar] / Unload threshold *)
    tLoadMin : TIME := T#30S;                (* 加载最小驻留，域 > T#0S [ms] / Minimum load dwell *)
    tUnloadMax: TIME := T#10M;               (* 卸载超时，域 > T#0S [ms] / Unload timeout *)
    tScan    : TIME := T#100MS;              (* 扫描周期，域 > T#0S [ms] / Scan period *)
    bEnable  : BOOL := TRUE;                 (* 使能 [-] / Enable *)
    bReset   : BOOL := FALSE;                (* 复位命令，上升沿清故障与告警 [-] / Reset command *)
END_VAR
VAR_OUTPUT
    bLoadCmd : BOOL;                         (* 加载命令信号 [-] / Load command *)
    bUnloadCmd: BOOL;                        (* 卸载命令信号 [-] / Unload command *)
    bMaintWarn: BOOL;                        (* 维护级告警锁存（卸载超时，复位沿清，边界③）[-] / Maintenance warning latched *)
    bSensorBad: BOOL;                        (* 压力传感器失效当拍出口（边界⑤）[-] / Sensor bad outlet *)
    eState   : E_DL_AclState;                (* 状态出口 / State outlet *)
    eCause   : E_DL_AclCause;                (* 成因出口（R190 归因唯一） / Cause outlet *)
    bError   : BOOL;                         (* 故障锁存标志 [-] / Fault latch flag *)
END_VAR
VAR
    _eState : E_DL_AclState := E_DL_AclState.eIdle;  (* 内部相位（CASE 唯一写入目标） / Internal phase *)
    _eCause : E_DL_AclCause := E_DL_AclCause.eNone;  (* 成因锁存量 / Latched cause *)
    rtReset : R_TRIG;                        (* 复位沿实例，段 0 无条件调用 / Reset edge instance *)
    tonLoad : TON;                           (* 加载驻留计时（IN 串 eLoad 相闸，R40） / Load dwell timer *)
    tonUnl  : TON;                           (* 卸载持续计时（IN 串 eUnload 相闸，R40） / Unload duration timer *)
    _bFault : BOOL;                          (* 故障锁存位 / Latched fault bit *)
    _bCfgBad: BOOL;                          (* 组态非法当拍量 / Illegal config this scan *)
    _bFin   : BOOL;                          (* 压力有限性当拍量（边界⑤） / Pressure finiteness *)
    _bUnlReq: BOOL;                          (* 卸载请求暂存量（驻留期内不丢，边界④） / Buffered unload request *)
    _fDtSec : REAL;                          (* 扫描周期秒值（信息级备用派生）[s] / Scan period seconds *)
END_VAR
VAR CONSTANT
    DL_ACL_EPS : REAL := 1.0E-6;             (* 判零容差 [-] / Epsilon *)
END_VAR

(* —— 段 0：当拍判据派生 + 实例无条件刷新（R228A；TON 全段 0 无 IF 包裹，R40） —— *)
_bCfgBad := NOT (fLoadTh < fUnloadTh)                    (* 压力带组态闸：加载阈 < 卸载阈（边界①） / Band config gate *)
            OR (fLoadTh <= DL_ACL_EPS)                   (* 加载阈正域闸 / Load threshold gate *)
            OR NOT (tLoadMin > T#0S) OR NOT (tUnloadMax > T#0S) OR NOT (tScan > T#0S);   (* 周期域闸 / Period gates *)
rtReset(CLK := bReset);                                  (* 复位沿每拍必调 / Reset edge every scan *)
_bFin := (fPress = fPress) AND ((fPress - fPress) = (fPress - fPress));   (* 压力 NaN 自反 + Inf 差判闸（边界⑤） / Pressure NaN and Inf gate *)
_fDtSec := TIME_TO_LREAL(tScan) / 1000.0;                (* 扫描周期秒化（除子常量 1000） / Scan period seconds *)
tonLoad(IN := (_eState = E_DL_AclState.eLoad), PT := tLoadMin);          (* 加载驻留：相位闸 + 无条件调用（R40） / Load dwell timer *)
tonUnl(IN := (_eState = E_DL_AclState.eUnload), PT := tUnloadMax);       (* 卸载持续：相位闸 + 无条件调用（R40） / Unload timer *)

(* —— 段 1：单拍量预清零（R107） —— *)
bLoadCmd := FALSE;                                       (* 加载命令出口预清（派生拍覆盖） / Load command preset *)
bUnloadCmd := FALSE;                                     (* 卸载命令出口预清 / Unload command preset *)
bSensorBad := FALSE;                                     (* 传感器失效当拍出口预清 / Sensor bad preset *)

(* —— 段 2：复位沿处理（作用域：清故障 + 清维护告警 + 迁 eIdle，R283 逐项声明） —— *)
IF rtReset.Q THEN
    _bFault := FALSE;                                    (* 清故障锁存 / Clear fault *)
    _eCause := E_DL_AclCause.eNone;                      (* 清成因 / Clear cause *)
    bMaintWarn := FALSE;                                 (* 清维护告警锁存 / Clear maintenance warning *)
    _bUnlReq := FALSE;                                   (* 清卸载请求暂存 / Clear buffered request *)
    _eState := E_DL_AclState.eIdle;                      (* 迁未使能相 / Back to idle *)
END_IF

(* —— 段 3：组态故障锁存（锁存至复位沿，R189） —— *)
IF _bCfgBad AND NOT _bFault THEN
    _bFault := TRUE;                                     (* 锁存故障位 / Latch fault *)
    _eCause := E_DL_AclCause.eCfgIllegal;                (* 成因：组态非法 / Cause illegal config *)
    _eState := E_DL_AclState.eFault;                     (* 同步迁故障相 / Migrate to fault *)
END_IF

(* —— 段 4：CASE 主状态机（ELSE 兜底迁 eFault，红线 6） —— *)
CASE _eState OF
    E_DL_AclState.eIdle:                                 (* 未使能：命令全停确定值 / Idle *)
        bLoadCmd := FALSE;                               (* 失能加载命令 FALSE / Disabled load false *)
        bUnloadCmd := FALSE;                             (* 失能卸载命令 FALSE / Disabled unload false *)
        IF bEnable AND NOT _bFault THEN
            _eState := E_DL_AclState.eLoad;              (* 使能先入加载相（建压优先） / Enter loading *)
        END_IF
    E_DL_AclState.eLoad:                                 (* 加载相：驻留 + 双阈迟滞切换 / Loading *)
        IF NOT bEnable THEN
            _eState := E_DL_AclState.eIdle;              (* 失能回未使能 / Back to idle *)
        ELSIF NOT _bFin THEN
            bSensorBad := TRUE;                          (* 传感器失效：保持当前态（边界⑤） / Sensor bad hold *)
        ELSE
            IF fPress >= fUnloadTh THEN
                _bUnlReq := TRUE;                        (* 驻留期内卸载请求暂存不丢（边界④） / Buffer unload request *)
            END_IF
            IF tonLoad.Q AND _bUnlReq THEN               (* 驻留满 + 有暂存请求：迁卸载（边界④） / Dwell done and request *)
                _bUnlReq := FALSE;                       (* 请求消费清零 / Request consumed *)
                _eState := E_DL_AclState.eUnload;        (* 迁卸载相 / To unloading *)
            END_IF
        END_IF
    E_DL_AclState.eUnload:                               (* 卸载相：下阈回加载 + 超时维护告警 / Unloading *)
        IF NOT bEnable THEN
            _eState := E_DL_AclState.eIdle;              (* 失能回未使能 / Back to idle *)
        ELSIF NOT _bFin THEN
            bSensorBad := TRUE;                          (* 传感器失效：保持当前态（边界⑤） / Sensor bad hold *)
        ELSE
            IF tonUnl.Q THEN                             (* 卸载持续超时（边界③） / Unload timeout *)
                bMaintWarn := TRUE;                      (* 维护级告警锁存（复位沿清，不自动停机） / Maintenance warning latch *)
                _eCause := E_DL_AclCause.eUnloadTime;    (* 成因：卸载超时（信息级不置 bError，边界③） / Cause unload time *)
            END_IF
            IF fPress <= fLoadTh THEN                    (* 压力回落到加载阈：迁加载（双阈迟滞直比，边界②） / Back to load *)
                _eState := E_DL_AclState.eLoad;          (* 迁加载相 / To loading *)
            END_IF
        END_IF
    E_DL_AclState.eFault:                                (* 故障相：命令全停冻结，仅复位沿出 / Fault *)
        ;                                                (* 锁存回放（R28） / Replay from latch *)
    ELSE                                                 (* 非法相位兜底迁安全态 / Illegal phase fallback *)
        _eState := E_DL_AclState.eFault; _bFault := TRUE;    (* 迁故障相 + 同步锁存 / To fault and latch *)
        _eCause := E_DL_AclCause.ePhaseBad;              (* 成因：非法相位 / Cause illegal phase *)
END_CASE

(* —— 段 5：出口映射（名实双出口，R191；bError/eState 同源） —— *)
bLoadCmd := (_eState = E_DL_AclState.eLoad);             (* 加载命令 = 加载相镜像 / Load command mirror *)
bUnloadCmd := (_eState = E_DL_AclState.eUnload);         (* 卸载命令 = 卸载相镜像 / Unload command mirror *)
bError := _bFault;                                       (* 故障标志镜像 / Fault flag mirror *)
eState := _eState;                                       (* 状态出口 / State outlet *)
eCause := _eCause;                                       (* 成因出口 / Cause outlet *)
END_FUNCTION_BLOCK

(* ---- FB_DL_AirDryerDiag.st ---- *)
(*
  ==================================================================
  组件名 Component  : FB_DL_AirDryerDiag
  分类   Category   : DL_Device
  前缀   Naming     : FB_DL_ ｜ b/n/u/f/t/e/st 类型前缀制（R265）
  复杂度 Complexity  : 中
  版本   Version    : 1.0.0
  功能   Purpose    : 压缩空气干燥机诊断（露点越限 + 再生阀时序状态机 + 切换周期劣化档）。
  来源   Source     : t2-2-lbp（干燥机诊断公开工艺语义）
  平台   Platform   : 纯 IEC 61131-3（TON / R_TRIG / CASE / TIME_TO_DINT），三平台通用
  分工声明 Split     : 与 FB_DL_DryerProtect（停机保护属主，若在册）分工——本件
                      只做诊断与周期劣化分档，不做停机联锁（R216 双向互引）。
  作者   Author     : 道莅代码库 · PLC 编程专家（R61）
  归属 Ownership     : E_DL_DryerPhase 属主为本文件（全库唯一定义，R264）；
                      引用件只引用不重声明。
  ------------------------------------------------------------------
  边界 Boundary     :
                      一 露点非有限闸逐个点名（R272：fDewPnt / fDewLim /
                         fDeg1Ratio / fDeg2Ratio 四个浮点引脚逐个判）；
                      二 再生切换周期劣化分档阈值全提为输入（fDeg1Ratio /
                         fDeg2Ratio [-]，实测周期与名义周期之比阈值，R 红线 7）；
                         组态递增配比违反判组态锁存（070F）；
                      三 状态机 CASE 必带 ELSE 兜底（R25 批次教训）；TON /
                         R_TRIG 段 0 无条件刷新（禁入分支，R7）；
                      四 故障锁存解除式逐条自证：bReset 上升沿清四锁存（恒可达，
                         R152 自证）；出口锁存回放优先（R187）；
                      五 周期换算：TIME 经 TIME_TO_DINT 落毫秒再升 LREAL 比
                         值（除零由组态闸 tCycleNom > 0 前置证明）；
                      六 无全局、无外部变量、无物理地址。
  错误码   Codes    :
    16#0003_070B【故障级】露点越限（fDewPnt > fDewLim），锁存至复位沿
    16#0003_070C【故障级】再生切换周期劣化二档（比值 ≥ fDeg2Ratio），锁存至复位沿
    16#0003_070D【故障级】露点入参非有限，锁存至复位沿
    16#0003_070E【信息级】再生切换周期劣化一档（比值 ≥ fDeg1Ratio，逐拍重算）
    16#0003_070F【故障级】组态非法（比值阈递增违反或名义周期 ≤ 0），锁存至复位沿
  验收   Acceptance :
    算法已证（脚本）：未跑 ｜ 编译器已证（三平台）：未跑
    V1 露点 -40、限 -20 → 无故障；V2 露点 -15 → 码 070B 锁存
    V3 实测周期 2 倍名义（阈 1.8）→ 码 070C 锁存；1.5 倍 → 070E 信息级
  修订记录 Revision  :
    2026-11-21  v1.0.0  R61 首版（批 4 · 序号 14）
  ==================================================================
*)
TYPE E_DL_DryerPhase :
(
    eDrying := 0,  // 吸附相：干燥塔在工作 / the drying phase, the tower working
    eRegen  := 10, // 再生相：再生阀开 / the regeneration phase, the valve open
    eFault  := 20  // 故障相：锁存待复位 / the fault phase latched until the reset
);
END_TYPE

FUNCTION_BLOCK FB_DL_AirDryerDiag
VAR_INPUT
    bEnable     : BOOL := TRUE;   // 使能，FALSE 时冻结诊断出口（R191 声明行）/ the enable, false freezes the diagnosis outlet
    bReset      : BOOL := FALSE;  // 故障复位电平，上升沿清锁存 / the fault reset level
    bRegenValve : BOOL := FALSE;  // 再生阀开反馈电平 [-] / the regeneration valve open feedback
    fDewPnt     : LREAL := -40.0; // 露点实测值 [摄氏度] / the measured dew point
    fDewLim     : LREAL := -20.0; // 露点上限 [摄氏度] / the dew point limit
    tCycleNom   : TIME := T#6H;   // 名义再生切换周期 [毫秒] / the nominal switch cycle
    fDeg1Ratio  : LREAL := 1.3;   // 劣化一档比值阈 [-] / the degradation level one ratio threshold
    fDeg2Ratio  : LREAL := 1.8;   // 劣化二档比值阈 [-] / the degradation level two ratio threshold
END_VAR
VAR_OUTPUT
    eState     : E_DL_DryerPhase;       // 主状态机当前态 [状态] / the current state
    bDewHigh   : BOOL := FALSE;         // 露点越限锁存指示 [-] / the dew over limit latched indicator
    bDeg1      : BOOL := FALSE;         // 劣化一档指示（信息级逐拍）[-] / the degradation level one indicator
    bDeg2      : BOOL := FALSE;         // 劣化二档锁存指示 [-] / the degradation level two latched indicator
    bError     : BOOL := FALSE;         // 故障锁存位（与锁存同源，R191）/ the fault bit from the latch
    bValid     : BOOL := FALSE;         // 诊断可用标志 [-] / the diagnosis usable flag
    eErr       : UDINT := 16#0000_0000; // 错误码，0 = 正常 / the error code, zero is ok
END_VAR
VAR
    _bInit     : BOOL := FALSE; // 首拍初始化标志（R310）/ the first scan flag
    _eState    : E_DL_DryerPhase := E_DL_DryerPhase.eDrying; // 内部状态寄存器 / the internal state register
    _bDewFlt   : BOOL := FALSE; // 露点越限锁存副本 / the dew fault latch copy
    _bDeg2Flt  : BOOL := FALSE; // 劣化二档锁存副本 / the level two latch copy
    _bDewNF    : BOOL := FALSE; // 露点非有限锁存副本 / the dew non finite latch copy
    _bCfgBad   : BOOL := FALSE; // 组态非法锁存副本 / the configuration latch copy
    _bFin      : BOOL := FALSE; // 四浮点引脚非有限闸结果（逐拍重算）/ the finiteness gate result
    _fRatio    : LREAL := 0.0;  // 实测周期与名义周期比 [-] / the measured to nominal ratio
    _tNomMs    : LREAL := 0.0;  // 名义周期 [毫秒] / the nominal cycle in milliseconds
    _tMeasMs   : LREAL := 0.0;  // 上一周实测周期 [毫秒] / the last measured cycle in milliseconds
    _tPrvSnap  : TIME := T#0S;  // 上拍周期计时快照（R 实战规则 1②）/ the previous cycle timing snapshot
    rtValve    : R_TRIG; // 再生阀开沿实例，段 0 无条件刷新 / the valve open edge instance
    rtReset    : R_TRIG; // 复位沿实例，段 0 无条件刷新 / the reset edge instance
    tonCycle   : TON;    // 切换周期实测计时器，段 0 无条件刷新 / the cycle measurement timer
END_VAR

// 段 0｜定时器与沿检测无条件周期刷新（禁入分支，R7）/ segment 0, the unconditional refresh
rtValve(CLK := bRegenValve); // 再生阀开沿 / the valve open edge
rtReset(CLK := bReset); // 复位沿 / the reset edge
tonCycle(IN := bRegenValve, PT := tCycleNom); // 周期实测（阀开时长累计）/ the cycle timing during the valve open
IF rtValve.Q THEN // 新一周开始：锁存上一周时长快照（周界沿取快照）/ a new cycle latches the last duration snapshot
    _tPrvSnap := tonCycle.ET; // 上周时长快照 / the last duration snapshot
END_IF

// 段 1｜首拍初始化与复位沿作用域（R310 / R311）/ segment 1, the first scan init and the reset scope
IF NOT _bInit THEN // 首拍一拍 / the first scan
    _bInit := TRUE; // 置首拍标志 / raise the first scan flag
    _bDewFlt := FALSE; // 露点锁存显式清零 / clear the dew latch explicitly
    _bDeg2Flt := FALSE; // 劣化二档锁存显式清零 / clear the level two latch explicitly
    _bDewNF := FALSE; // 非有限锁存显式清零 / clear the non finite latch explicitly
    _bCfgBad := FALSE; // 组态锁存显式清零 / clear the configuration latch explicitly
    _eState := E_DL_DryerPhase.eDrying; // 状态显式落吸附相 / place the state to drying
END_IF
IF rtReset.Q THEN // 复位沿（作用域：清四锁存 + 迁相位，R311 声明）/ the reset edge with the declared scope
    _bDewFlt := FALSE; // 清露点锁存（解除路径：复位沿恒可达，R152 自证）/ clear the dew latch
    _bDeg2Flt := FALSE; // 清劣化二档锁存 / clear the level two latch
    _bDewNF := FALSE; // 清非有限锁存 / clear the non finite latch
    _bCfgBad := FALSE; // 清组态锁存 / clear the configuration latch
    _eState := E_DL_DryerPhase.eDrying; // 迁回吸附相 / back to drying
END_IF

// 段 2｜非有限闸与组态闸（R272 全量点名，边界一二）/ segment 2, the finiteness and the configuration gates
_bFin := (fDewPnt = fDewPnt) AND ((fDewPnt - fDewPnt) = (fDewPnt - fDewPnt))
AND (fDewLim = fDewLim) AND ((fDewLim - fDewLim) = (fDewLim - fDewLim))
AND (fDeg1Ratio = fDeg1Ratio) AND ((fDeg1Ratio - fDeg1Ratio) = (fDeg1Ratio - fDeg1Ratio))
AND (fDeg2Ratio = fDeg2Ratio) AND ((fDeg2Ratio - fDeg2Ratio) = (fDeg2Ratio - fDeg2Ratio)); // 四浮点引脚逐个自反 + 差值判 / the four floating pins tested one by one
IF NOT _bFin THEN // 入参非有限（露点成因独立锁存，R190）/ a non finite input latches the dew cause
    _bDewNF := TRUE; // 锁存非有限（070D）/ latch the non finite cause
END_IF
IF (fDeg1Ratio <= 1.0) OR (fDeg2Ratio <= fDeg1Ratio) OR (tCycleNom <= T#0S) THEN // 组态递增配比违反（边界二）/ the configuration monotone ratio violated
    _bCfgBad := TRUE; // 锁存组态非法（070F）/ latch the configuration fault
END_IF
_tNomMs := DINT_TO_LREAL(TIME_TO_DINT(tCycleNom)); // 名义周期毫秒化（TIME 口径，边界五）/ the nominal cycle in milliseconds

// 段 3｜露点越限判据（有限才判）/ segment 3, the dew over limit criterion
IF _bFin AND (fDewPnt > fDewLim) THEN // 露点越限（070B 独立成因）/ the dew over the limit
    _bDewFlt := TRUE; // 独立锁存 / latch the dew cause
END_IF

// 段 4｜周期比与劣化分档（周界沿快照换算，除零前置证明）/ segment 4, the cycle ratio and the degradation grades
IF rtValve.Q THEN // 新周界沿：换算上周比值 / a new cycle edge converts the last ratio
    _tMeasMs := DINT_TO_LREAL(TIME_TO_DINT(_tPrvSnap)); // 上周时长毫秒化 / the last duration in milliseconds
    IF _tNomMs > 0.0 THEN // 除零防护（组态闸已证 > 0，双保险）/ the division guard doubled
        _fRatio := _tMeasMs / _tNomMs; // 周期比（除子已证 > 0）/ the cycle ratio with a proven divisor
        IF _fRatio >= fDeg2Ratio THEN // 二档劣化（070C 独立成因）/ the level two degradation
            _bDeg2Flt := TRUE; // 独立锁存 / latch the level two cause
        END_IF
    END_IF
END_IF

// 段 5｜主状态机（ENUM + CASE，ELSE 兜底，边界三）/ segment 5, the main machine with the ELSE guard
CASE _eState OF
    E_DL_DryerPhase.eDrying: // 吸附相 / the drying phase
        IF bRegenValve THEN // 阀开反馈迁入再生相 / the valve open feedback migrates to regen
            _eState := E_DL_DryerPhase.eRegen; // 迁入再生相 / enter the regen phase
        ELSIF _bDewFlt OR _bDeg2Flt OR _bDewNF OR _bCfgBad THEN // 故障迁移（锁存复检，R274）/ the fault migration with the latch recheck
            _eState := E_DL_DryerPhase.eFault; // 迁入故障相 / enter the fault phase
        END_IF
    E_DL_DryerPhase.eRegen: // 再生相 / the regen phase
        IF NOT bRegenValve THEN // 阀关反馈迁回吸附相 / the valve closed feedback back to drying
            _eState := E_DL_DryerPhase.eDrying; // 迁回吸附相 / back to drying
        ELSIF _bDewFlt OR _bDeg2Flt OR _bDewNF OR _bCfgBad THEN // 故障迁移 / the fault migration
            _eState := E_DL_DryerPhase.eFault; // 迁入故障相 / enter the fault phase
        END_IF
    E_DL_DryerPhase.eFault: // 故障相：等复位沿（解除可达，边界四）/ the fault phase until the reset
        IF NOT (_bDewFlt OR _bDeg2Flt OR _bDewNF OR _bCfgBad) THEN // 四锁存已清才迁出（防清锁同拍重锁，FB50-1）/ the exit after all latches cleared
            _eState := E_DL_DryerPhase.eDrying; // 迁回吸附相 / back to drying
        END_IF
    ELSE // 非法枚举值拦截（兜底码走组态成因回放）/ the illegal enumeration guard
        _eState := E_DL_DryerPhase.eFault; // 落入故障相 / force to the fault phase
        _bCfgBad := TRUE; // 置锁存（ELSE 兜底码走组态成因回放）/ latch the configuration cause
END_CASE

// 段 6｜统一出口（锁存同源映射；一档信息级逐拍重算，R285）/ segment 6, the unified outlet
eState := _eState; // 状态出口 / the state outlet
bDewHigh := _bDewFlt; // 露点越限出口 / the dew outlet
bDeg2 := _bDeg2Flt; // 二档出口 / the level two outlet
bDeg1 := (NOT _bDeg2Flt) AND (_fRatio >= fDeg1Ratio); // 一档指示（逐拍重算，信息级不置 bError）/ the level one indicator recomputed
bError := _bDewFlt OR _bDeg2Flt OR _bDewNF OR _bCfgBad; // 故障位出口 / the fault bit outlet
bValid := (NOT bError) AND bEnable; // 诊断可用标志 / the usable flag
IF _bCfgBad THEN // 组态成因回放优先 / the configuration cause replays first
    eErr := 16#0003_070F; // 故障级：组态非法 / fault grade, the illegal configuration
ELSIF _bDewNF THEN // 非有限成因 / the non finite cause
    eErr := 16#0003_070D; // 故障级：露点入参非有限 / fault grade, the non finite dew input
ELSIF _bDewFlt THEN // 露点越限成因 / the dew cause
    eErr := 16#0003_070B; // 故障级：露点越限 / fault grade, the dew over the limit
ELSIF _bDeg2Flt THEN // 二档成因 / the level two cause
    eErr := 16#0003_070C; // 故障级：切换周期劣化二档 / fault grade, the cycle degradation level two
ELSE // 无故障 / no fault
    eErr := 16#0000_0000; // 正常 / ok
END_IF
END_FUNCTION_BLOCK

(* ---- FB_DL_AnalogDriftWatch.st ---- *)
(*
    FB_DL_AnalogDriftWatch —— 模拟量双通道冗余漂移监测
    ------------------------------------------------------------------
    分类      : DL_Device / AnalogHealth
    前缀      : FB_DL_
    版本      : 1.0.0
    溯源      : clean-room 自有实现；仅借鉴「双通道偏差指数遗忘累积」的公开
                滤波/监测常识语义，未复制任何闭源厂商源码，码位 100% 自有
    平台      : 纯 IEC 61131-3，CODESYS V3.5+ / TwinCAT 3 / InoProShop / Machine Expert 通用
    作者      : 道莅代码库 · PLC编程专家（R76 冲刺批 C3 · #4）
    ------------------------------------------------------------------
    功能说明  : 双通道模拟量 fValA/fValB 冗余漂移监测：偏差 |fValA - fValB| 按指数
                遗忘累积为漂移估计 fDrift（α = fDtSec / (fTauSec + fDtSec)，分母
                门禁防除零，α 天然落在 (0,1] 无需再钳位）。漂移超 fWarnTh 报预警
                （bWarn，信息/预警级，不置 bError）；超 fFaultTh 报故障并判主通道
                失可信（bATrust = FALSE），锁存至 bReset 复位沿。任一通道非有限值
                （NaN f<>f、±Inf (f-f)<>(f-f)）按「单边失可信」处理：该通道信任
                标志置 FALSE、漂移估计冻结不更新、条件级故障码每拍重发布，
                不误报漂移，条件消失自动恢复。
                边界：只产出漂移估计与信任判定，不做通道切换、不修正采样值。
    错误码    : 16#0005_2000 参数非法（时间常数/周期非正或非有限 / 阈值非正 /
                             fFaultTh <= fWarnTh）——故障级，锁存至复位沿
                16#0005_2001 漂移估计超故障阈值，主通道 A 判失可信——故障级，
                             锁存至 bReset 复位沿
                16#0005_2002 通道 A 非有限，单边失可信，估计冻结——条件级故障，
                             条件存在每拍重发布、条件消失自动恢复，不锁存
                16#0005_2003 通道 B 非有限，单边失可信，估计冻结——条件级故障，
                             同 2002 口径
                16#0005_2004 漂移估计超预警阈值——预警级，超阈期间持续发布，不置 bError
                16#0005_2005 CASE 落 ELSE 兜底——故障级，锁存至复位沿
    码位总账  : 16#0005_2000..2005 全部定义并使用，无空悬码位
    状态机    : E_DL_DriftState（eIdle / eRun / eFault），CASE 含 ELSE 兜底：落 ELSE
                置 16#0005_2005 并回 eFault。eIdle 时不背书：bATrust/bBTrust 置
                FALSE（监测未运行不给可信结论）；eFault 锁存码回放，bReset 上升沿
                且参数已合法时清零漂移估计回 eIdle。
    定时器    : 本件无 TON；仅一只 R_TRIG 在本体段 1 无条件周期刷新（R7）。
    防御口径  : α 分母 (fTauSec + fDtSec) 强制 > 0 且两参非有限门禁后才做除法，
                绝无除零；阈值比较用严格大于（禁 =/<>）；漂移估计仅当双通道
                均有限时更新，冻结路径不触碰累计量。
    修订记录  : 2026-11-23 v1.0.0 首次入库（R76 冲刺批 C3 · #4）
*)
TYPE E_DL_DriftState :
(
    eIdle  := 0,   // 待机，监测未投运，不背书信任标志 / idle, monitoring off, trust flags not endorsed
    eRun   := 10,  // 运行，每拍更新漂移估计并判阈 / running, drift estimate updated and thresholds judged every scan
    eFault := 20   // 故障，锁存码回放，主通道判失可信 / fault, latch replayed, the main channel is distrusted
);
END_TYPE

FUNCTION_BLOCK FB_DL_AnalogDriftWatch
VAR_INPUT
    fValA    : LREAL;                  // 主通道 A 采样值 [工程单位] / main channel A sample [engineering unit]
    fValB    : LREAL;                  // 备通道 B 采样值 [工程单位] / redundant channel B sample [engineering unit]
    fWarnTh  : LREAL := 1.0;           // 漂移预警阈值 [工程单位]，必须大于 0 / drift warning threshold [engineering unit], must exceed zero
    fFaultTh : LREAL := 2.0;           // 漂移故障阈值 [工程单位]，必须大于 fWarnTh / drift fault threshold, must exceed fWarnTh
    fTauSec  : LREAL := 5.0;           // 指数遗忘时间常数 [s]，必须大于 0 / exponential forgetting time constant [s], must exceed zero
    fDtSec   : LREAL := 0.1;           // 采样周期 [s]，必须大于 0 / sampling period [s], must exceed zero
    bMonEn   : BOOL := TRUE;           // 监测投运命令 / monitoring enable command
    bReset   : BOOL;                   // 故障复位请求，上升沿生效 / fault reset request, edge-active
END_VAR
VAR_OUTPUT
    fDrift   : LREAL;                  // 漂移估计 [工程单位]，仅双通道有限时更新 / drift estimate [engineering unit], updated only when both channels are finite
    bWarn    : BOOL;                   // 预警标志，超 fWarnTh 置位 / warning flag, raised above fWarnTh
    bATrust  : BOOL;                   // 主通道 A 可信标志，非有限或漂移故障置 FALSE / main channel trust flag, FALSE when non-finite or on a drift fault
    bBTrust  : BOOL;                   // 备通道 B 可信标志，非有限置 FALSE / redundant channel trust flag, FALSE when non-finite
    eState   : E_DL_DriftState;        // 当前状态镜像输出 / current state mirror output
    nErrCode : UDINT;                  // 错误码，0 = 无错；锁存级回放、条件级随条件发布 / error code, 0 = none; latched codes replayed, conditional codes per condition
    bError   : BOOL;                   // 故障级标志，仅故障级码置位 / fault-class flag, raised only by fault-class codes
    bValid   : BOOL;                   // 输出可用标志，= NOT bError / outputs valid flag, equals NOT bError
END_VAR
VAR
    _eState    : E_DL_DriftState;      // 当前状态 / current state
    _uErrLatch : UDINT;                // 锁存故障码副本（2000/2001/2005），故障态每拍回放 / latched fault code replayed inside the fault state
    rtReset    : R_TRIG;               // 复位上升沿检测 / reset rising-edge detector
    _fAlpha    : LREAL;                // 遗忘系数 α = fDtSec/(fTauSec+fDtSec)，(0,1] / forgetting factor within (0,1]
    _fDiff     : LREAL;                // 本拍双通道偏差绝对值 [工程单位] / absolute inter-channel deviation this scan
    _bAOk      : BOOL;                 // 通道 A 有限标志 / channel A finite flag
    _bBOk      : BOOL;                 // 通道 B 有限标志 / channel B finite flag
    _bParOk    : BOOL;                 // 参数门禁结果 / parameter gate result
END_VAR
VAR CONSTANT
    DL_ADW_ONE  : LREAL := 1.0;        // 遗忘权重基值 [无量纲] / forgetting weight base [dimensionless]
    DL_ADW_ZERO : LREAL := 0.0;        // 零值常量，避免裸字面量 [工程单位] / zero constant avoiding a bare literal [engineering unit]
END_VAR

// 段 1｜边缘检测无条件周期刷新（R7：严禁放入 IF / CASE；本件无 TON）
// segment 1, edge detector refreshed unconditionally, never inside IF/CASE; no TON in this FB
rtReset(CLK := bReset);

// 段 2｜输出与错误状态预置；锁存级故障态从锁存副本回放（R45 配对）
// segment 2, preset outputs and error status; latched fault states replay from the latch
bWarn := FALSE;                        // 预置无预警 / preset no warning
bATrust := TRUE;                       // 预置主通道可信 / preset main channel trusted
bBTrust := TRUE;                       // 预装备通道可信 / preset redundant channel trusted
nErrCode := 0;                         // 预置无错误码 / preset no error code
bError := FALSE;                       // 预置无故障标志 / preset no fault flag
bValid := TRUE;                        // 预置输出可用 / preset outputs valid
IF _eState = E_DL_DriftState.eFault THEN
    nErrCode := _uErrLatch;            // 重发布锁存故障码，HMI 不会看到码位闪断 / republish the latched fault code
    bError := TRUE;                    // 故障态恒置故障标志 / fault flag stays raised in the fault state
    bValid := FALSE;                   // 故障态输出不可信 / outputs not valid in the fault state
    IF _uErrLatch = 16#0005_2001 THEN
        bATrust := FALSE;              // 漂移故障回放期主通道持续失可信 / main channel stays distrusted while the drift fault replays
    END_IF
END_IF

// 段 3｜通道有限判定 + α 防除零计算：非有限按单边失可信口径，α 仅在门禁通过后计算
// segment 3, per-channel finite test and the divide-guarded alpha; non-finite follows the single-side distrust policy
_bAOk := NOT ((fValA <> fValA) OR ((fValA - fValA) <> (fValA - fValA)));  // A 非有限判定（NaN 自不等 / Inf 自差不等）/ A NaN via self-inequality, Inf via self-difference
_bBOk := NOT ((fValB <> fValB) OR ((fValB - fValB) <> (fValB - fValB)));  // B 非有限判定，口径同 A / channel B tested the same way
_bParOk := (fTauSec > DL_ADW_ZERO) AND (fDtSec > DL_ADW_ZERO)
       AND (fWarnTh > DL_ADW_ZERO) AND (fFaultTh > fWarnTh)
       AND NOT ((fTauSec <> fTauSec) OR ((fTauSec - fTauSec) <> (fTauSec - fTauSec)))
       AND NOT ((fDtSec <> fDtSec) OR ((fDtSec - fDtSec) <> (fDtSec - fDtSec)))
       AND NOT ((fWarnTh <> fWarnTh) OR ((fWarnTh - fWarnTh) <> (fWarnTh - fWarnTh)))
       AND NOT ((fFaultTh <> fFaultTh) OR ((fFaultTh - fFaultTh) <> (fFaultTh - fFaultTh)));
IF _bParOk THEN
    _fAlpha := fDtSec / (fTauSec + fDtSec); // 分母 = fTauSec + fDtSec > fDtSec > 0，绝无除零；α 天然 (0,1] / denominator exceeds fDtSec, no zero division, alpha within (0,1]
END_IF
IF (NOT _bParOk) AND (_eState <> E_DL_DriftState.eFault) THEN
    _uErrLatch := 16#0005_2000;        // 锁存参数非法码 / latch the illegal parameter code
    nErrCode := 16#0005_2000;          // 故障级码赋值 3 行内置 bError / fault-class assignment with bError inline
    bError := TRUE;
    bValid := FALSE;
    _eState := E_DL_DriftState.eFault; // 参数不可信直接转故障 / untrusted parameters jump to fault
END_IF

// 段 4｜主状态机：CASE + ELSE 兜底（R6）；漂移更新仅在 eRun 且双通道有限时执行
// segment 4, main state machine, CASE with ELSE fallback; the drift update runs only in eRun with both channels finite
CASE _eState OF
E_DL_DriftState.eIdle:
    // 拍 N 进入：复位后或未投运；本拍行为：不背书信任标志、估计保持清零；拍 N+1 转出：投运且参数合法 → eRun
    // entered after reset or when disabled; no trust endorsement and the estimate stays cleared; exits to eRun on enable with legal parameters
    bATrust := FALSE;                  // 监测未运行不给可信结论 / no trust verdict while monitoring is off
    bBTrust := FALSE;                  // 备通道同样不背书 / the redundant channel is not endorsed either
    fDrift := DL_ADW_ZERO;             // 估计清零，防旧值带病入运行 / clear the estimate so no stale value carries over
    IF bMonEn AND _bParOk THEN
        _eState := E_DL_DriftState.eRun; // 进运行相 / enter the run phase
    END_IF

E_DL_DriftState.eRun:
    // 拍 N 进入：投运且参数合法；本拍行为：双通道有限则更新估计并判阈，单边非有限则
    // 冻结估计、发布条件级码；拍 N+1 转出：超故障阈 → eFault（2001）；参数门禁 → eFault（段 3）
    // entered on enable with legal parameters; the estimate updates and thresholds are judged when both channels
    // are finite, otherwise it freezes with a conditional code; exits to eFault above the fault threshold (2001)
    IF (NOT _bAOk) OR (NOT _bBOk) THEN
        // 单边失可信：估计冻结不更新，杜绝非有限值污染累计量（不误报漂移）
        // single-side distrust: freeze the estimate so non-finite values can never pollute the accumulator
        IF NOT _bAOk THEN
            bATrust := FALSE;              // 主通道失可信 / main channel distrusted
            nErrCode := 16#0005_2002;      // 条件级故障：条件存在每拍重发布、消失自动恢复 / conditional fault republished per scan
            bError := TRUE;                // 故障级码赋值 3 行内置 bError（条件级不锁存）/ fault-class trio, conditional not latched
            bValid := FALSE;
        END_IF
        IF NOT _bBOk THEN
            bBTrust := FALSE;              // 备通道失可信 / redundant channel distrusted
            nErrCode := 16#0005_2003;      // 双通道同拍非有限时 B 后赋值可见 / assigned after A so B wins when both fail together
            bError := TRUE;                // 故障级码赋值 3 行内置 bError / fault-class assignment with bError inline
            bValid := FALSE;
        END_IF
    ELSE
        _fDiff := ABS(fValA - fValB);      // 本拍偏差绝对值 [工程单位] / absolute deviation this scan
        fDrift := fDrift * (DL_ADW_ONE - _fAlpha) + _fDiff * _fAlpha; // 指数遗忘累积 / exponential forgetting accumulation
        IF fDrift > fFaultTh THEN
            _uErrLatch := 16#0005_2001;    // 锁存漂移故障码 / latch the drift fault code
            nErrCode := 16#0005_2001;      // 故障级码赋值 3 行内置 bError / fault-class assignment with bError inline
            bError := TRUE;
            bValid := FALSE;
            bATrust := FALSE;              // 主通道判失可信 / main channel distrusted
            _eState := E_DL_DriftState.eFault; // 转故障锁存 / go to fault and latch
        ELSIF fDrift > fWarnTh THEN
            bWarn := TRUE;                 // 预警置位 / raise the warning
            nErrCode := 16#0005_2004;      // 预警级：超阈期间持续发布，不置 bError / warning class, no fault flag
        END_IF
    END_IF

E_DL_DriftState.eFault:
    // 拍 N 进入：参数非法或漂移超故障阈；本拍行为：锁存码回放、信任标志按码维持；
    // 拍 N+1 转出：bReset 上升沿且参数已合法 → eIdle（估计清零重新起算）
    // entered on illegal parameters or a drift fault; the latch replays and trust follows the code;
    // exits to eIdle on a reset edge with legal parameters, the estimate restarts from zero
    IF rtReset.Q AND _bParOk THEN
        _uErrLatch := 0;                   // 清锁存码 / clear the latched code
        fDrift := DL_ADW_ZERO;             // 估计清零重新起算 / restart the estimate from zero
        _eState := E_DL_DriftState.eIdle;  // 回待机等投运 / back to idle awaiting enable
    END_IF

ELSE
    // 非法状态拦截：任何未定义枚举值一律锁存兜底码并转故障（R6）
    // illegal-state interception, any undefined enum value latches the fallback code and goes to fault
    _uErrLatch := 16#0005_2005;            // 锁存兜底码 / latch the fallback code
    nErrCode := 16#0005_2005;              // 故障级码赋值 3 行内置 bError / fault-class assignment with bError inline
    bError := TRUE;
    bValid := FALSE;
    _eState := E_DL_DriftState.eFault;
END_CASE

// 段 5｜状态镜像输出
// segment 5, state mirror output
eState := _eState;                     // 状态镜像输出 / state mirror output

END_FUNCTION_BLOCK

(* ---- FB_DL_AnalogOutFailsafe.st ---- *)
(*
  ==================================================================
  组件名 Component  : FB_DL_AnalogOutFailsafe
  分类   Category   : DL_Device
  前缀   Naming     : FB_DL_ ｜ b/n/u/f/t/e 类型前缀制（R265）
  版本   Version    : 1.0.1
  功能   Purpose    : 模拟量输出失保通道：正常相把 fOutReq（0~100 钳位）经
                      斜坡限速送达 fOutAct；看门狗超时 / 请求非有限 / 配置
                      非法任一成立即锁存故障，按 eFailMode 走冻结或安全值
                      侧（安全值侧斜坡回程限速，不跳变）。bError 锁存，
                      解除式（可达自证·电平式 v1.0.1）：使能 + 心跳在 +
                      无超时 + 配置恢复 + 请求有限 → 清锁存回正常相。
  来源   Source     : t2-8-ne43（NE43 失效安全方向口径：借「失效落安全侧」
                      语义，实现零源码复制）
  互引   Cross-ref  : FB_DL_AnalogSignalHealth（上游信号健康诊断件，可把其
                      bHealthy 布到本件 bWatchdog 心跳引脚）
  平台   Platform   : 纯 IEC 61131-3（TON/R_TRIG/ENUM+CASE/LREAL 四则）
  依赖   Depends    : 仅 Standard.library（TON/R_TRIG 属标准件）
  归属   Ownership  : E_DL_FailMode 与 E_DL_AnaOutFsState 属主为本文件
                      （全库唯一定义，R264）；引用件只引用不重声明。
  设计偏差 Deviation: 时间基准按本库「时间注入」纪律：新增输入 fCallCycleS
                      （调用方注入扫描周期 [s]，FB_DL_CycleTimeMeasure 语义），
                      本件不读平台时刻函数；斜坡步长 = fRampRatePctS × fCallCycleS。
  红线   Redline    : R1 零全局/VAR_EXTERNAL/R2 零 %I/%Q/R3 纯 IEC 标准
                      R4 输出 0~100 显式钳位 + 非有限三闸（请求/安全值/周期）
                      + 除法零处（无除法面）/R5 全变量双语同行注释
                      R6 ENUM+CASE 含 ELSE 兜底，eFault 分支显式出现
                      R7 tonWd 段 0 无条件刷新（IN = NOT bWatchdog，
                      v1.0.1 订正反相：断线达整定才超时）
                      R8 钳位与阈值常量化
  错误码 Codes      : 16#0007_1001【故障级·锁存】看门狗超时（心跳丢失）
                      16#0007_1002【故障级·锁存】配置非法（斜坡速率 ≤ 0 /
                      安全值非有限 / 扫描周期 ≤ 0）
                      16#0007_1003【故障级·锁存】请求非有限（NaN/±Inf）
                      锁存解除（可达自证·电平式 v1.0.1）：bEnable + 心跳在
                      （bWatchdog=TRUE 且 tonWd 未超时）+ 配置恢复 + 请求
                      有限 → 清锁存回 eNormal；三成因解除条件均为电平恒可
                      满足，无「置位即永久」路径（R66 终审修：弃沿式解除，
                      恒真心跳缺省组态下沿式对 1002/1003 不可达）。
  码位反证 Note     : 1001/1002/1003 分立依据（R190 归因唯一）：三成因
                      （超时/配置/请求）各有独立观测入口与独立处置面，
                      禁共用码导致某成因永不赋值。
  验收   Acceptance : V1 正常跟踪：斜坡达目标 + bAtCmd 语义 ｜ V2 心跳断
                      tWdTimeout → 锁存 1001 + 按 eFailMode 动作 ｜
                      V3 fOutReq=NaN → 锁存 1003 + 安全侧 ｜ V4 fRampRatePctS=0
                      → 锁存 1002 ｜ V5 故障中恢复心跳 + 使能 → 解锁回正常
                      ｜ V6 eFreeze → 冻结保持当前值不回程 ｜ V7 全程输出
                      不出 [0,100]
  变更   Revision   : 2026-11-22  v1.0.0  R66 首版（编码阶段批 3 序 7）
                      2026-11-22  v1.0.1  R66 终审就地修（3 严重）：①tonWd
                      IN 反相订正（IN=NOT bWatchdog，原写法健康心跳驻留
                      tWdTimeout 即误锁 1001、真断线反不检测）；②锁存期
                      eFrozen/eSafeHold 运行路径打通（段 6 弃整体旁路，段 5
                      改锁存起点单次迁入）；③锁存解除弃沿式改电平式（删
                      rtWdRecover，恒真心跳下沿式对 1002/1003 不可达）。
  ==================================================================
*)
TYPE E_DL_FailMode :
(
    eFreeze    := 0,  // 失保动作=冻结保持当前输出 [-] / the fail action freezes the current output
    eSafeValue := 1   // 失保动作=斜坡回程到 fSafeValue [-] / the fail action ramps to the safe value
);
END_TYPE

TYPE E_DL_AnaOutFsState :
(
    eIdle    := 0,   // 失能：bEnable=FALSE，输出冻结保持 [-] / the disabled phase, outputs frozen
    eNormal  := 10,  // 正常：斜坡跟踪请求 [-] / the normal phase, ramping toward the request
    eFrozen  := 20,  // 失保冻结：保持故障瞬间的当前值 [-] / the fail frozen phase, holding the fault time value
    eSafeHold:= 30,  // 失保安全值：斜坡回程到安全值并保持 [-] / the fail safe phase, ramping to the safe value
    eFault   := 40   // 锁存故障：锁存驻留，解除沿回正常 [-] / the latched fault phase dwelling until the release edge
);
END_TYPE

FUNCTION_BLOCK FB_DL_AnalogOutFailsafe
VAR_INPUT
    fOutReq      : LREAL := 0.0;    // 输出请求 [%]，0~100 钳位，非有限按安全侧 / the output request, clamped, non finite goes safe side
    bEnable      : BOOL := FALSE;   // 使能，FALSE 冻结输出保持（失能语义写死，FB33-4）[-] / the enable, false freezes the output
    bWatchdog    : BOOL := TRUE;    // 上游心跳电平（TRUE=心跳在）[-] / the upstream heartbeat level
    eFailMode    : E_DL_FailMode := E_DL_FailMode.eSafeValue; // 失保模式（冻结/安全值）[-] / the fail mode
    fSafeValue   : LREAL := 0.0;    // 失保安全值 [%]，须有限（非有限判配置非法）/ the fail safe value, must be finite
    fRampRatePctS: LREAL := 10.0;   // 斜坡速率 [%/s]，须 > 0（≤ 0 判配置非法）/ the ramp rate, must be positive
    tWdTimeout   : TIME := T#2S;    // 看门狗超时整定 [ms] / the watchdog timeout setting
    fCallCycleS  : LREAL := 0.01;   // 调用方注入扫描周期 [s]，须 > 0 / the caller injected scan cycle in seconds
END_VAR
VAR_OUTPUT
    fOutAct      : LREAL := 0.0;    // 实际输出 [%]，全程钳位 0~100 / the actual output, always clamped 0 to 100
    eState       : E_DL_AnaOutFsState := E_DL_AnaOutFsState.eIdle; // 状态机出口 [状态] / the state machine outlet
    bError       : BOOL := FALSE;   // 故障锁存标志（解除沿清除，R45 配对）/ the latched fault flag, cleared by the release edge
    uErrorId     : UDINT := 16#0000_0000; // 故障码，0=正常；锁存回放至解除沿 [码] / the latched fault code replayed to the release edge
END_VAR
VAR
    _bInit       : BOOL := FALSE;   // 首拍初始化标志（R310）/ the first scan flag
    _eState      : E_DL_AnaOutFsState := E_DL_AnaOutFsState.eIdle; // 内部状态寄存器 / the internal state register
    _bFaultLatch : BOOL := FALSE;   // 故障锁存副本（仅解除沿清除）/ the fault latch copy, cleared only by the release edge
    _uLatch      : UDINT := 16#0000_0000; // 故障码锁存副本（仅解除沿清除，FB33-1）/ the latched code copy
    _bCfgOk      : BOOL := FALSE;   // 本拍配置有效性 [-] / the per scan configuration validity
    _fStep       : LREAL := 0.0;    // 本拍斜坡步长 [%] / the per scan ramp step
    _fTarget     : LREAL := 0.0;    // 本拍斜坡目标 [%] / the per scan ramp target
    _bClampReq   : BOOL := FALSE;   // 本拍请求被钳位标志（信息性，未设码）[-] / the per scan request clamp flag, informational
    tonWd        : TON;             // 看门狗定时器实例，段 0 无条件刷新 / the watchdog timer instance refreshed unconditionally
END_VAR
VAR CONSTANT
    AOF_OUT_MIN  : LREAL := 0.0;      // 输出下限 [%] / the output lower clamp
    AOF_OUT_MAX  : LREAL := 100.0;    // 输出上限 [%] / the output upper clamp
    AOF_FIN_MAX  : LREAL := 1.7976931348623157E308; // LREAL 有限上限 / the finite LREAL limit
    AOF_ERR_NONE : UDINT := 16#0000_0000; // 无故障 [码] / no fault [code]
    AOF_ERR_WDTO : UDINT := 16#0007_1001; // 码 1001：看门狗超时 / code 1001, watchdog timeout
    AOF_ERR_CFG  : UDINT := 16#0007_1002; // 码 1002：配置非法 / code 1002, illegal configuration
    AOF_ERR_REQ  : UDINT := 16#0007_1003; // 码 1003：请求非有限 / code 1003, non finite request
END_VAR

(*------------------------------------------------------------------------------
 * 段 0｜定时器与沿检测无条件刷新区（红线 R7）：严禁移入 IF / CASE
 *      The timer and edge instances refresh unconditionally, never in a branch
 *-----------------------------------------------------------------------------*)
tonWd(IN := NOT bWatchdog, PT := tWdTimeout);   // 心跳断线计时（v1.0.1 订正 IN 反相：断线达整定才超时）/ the heartbeat loss timing, IN inverted per R66 review

(*------------------------------------------------------------------------------
 * 段 1｜首拍初始化：输出从钳位后的请求值起（避免首拍跳变）
 *      First scan init: the output starts from the clamped request
 *-----------------------------------------------------------------------------*)
IF NOT _bInit THEN
    _bInit := TRUE;                         // 首拍标志落位 / arm the first scan flag
    IF (fOutReq >= AOF_OUT_MIN) AND (fOutReq <= AOF_OUT_MAX) AND (fOutReq = fOutReq) THEN
        fOutAct := fOutReq;                 // 有限且在域内直接落位 / land directly when finite and inside
    ELSE
        fOutAct := AOF_OUT_MIN;             // 首拍非法请求落安全下限 / land on the safe lower limit
    END_IF
END_IF

(*------------------------------------------------------------------------------
 * 段 2｜配置闸（归因唯一 R190）：速率 ≤ 0 / 安全值非有限 / 周期 ≤ 0 → 配置非法
 *      The configuration gate with unique attribution per cause
 *-----------------------------------------------------------------------------*)
_bCfgOk := (fRampRatePctS > 0.0)
       AND (fSafeValue = fSafeValue) AND (ABS(fSafeValue) <= AOF_FIN_MAX)
       AND (fCallCycleS > 0.0) AND (fCallCycleS = fCallCycleS);   // 三配置面逐项闸 / each configuration face gated

(*------------------------------------------------------------------------------
 * 段 3｜故障成因判定与锁存（锁存回放，不在故障相按当下输入重推断）
 *      Fault cause determination and latching, replayed not re inferred in the fault phase
 *-----------------------------------------------------------------------------*)
IF tonWd.Q THEN                                // 成因一：心跳超时 / cause one, the heartbeat timeout
    _bFaultLatch := TRUE;
    _uLatch := AOF_ERR_WDTO;
ELSIF NOT _bCfgOk THEN                         // 成因二：配置非法 / cause two, illegal configuration
    _bFaultLatch := TRUE;
    _uLatch := AOF_ERR_CFG;
ELSIF (fOutReq <> fOutReq) OR (ABS(fOutReq) > AOF_FIN_MAX) THEN  // 成因三：请求非有限 / cause three, non finite request
    _bFaultLatch := TRUE;
    _uLatch := AOF_ERR_REQ;
END_IF

(*------------------------------------------------------------------------------
 * 段 4｜锁存解除（可达自证）：使能 + 无超时 + 配置恢复 + 心跳恢复上升沿
 *      The latch release, reachable by construction: enable, no timeout, config ok, heartbeat re entry edge
 *-----------------------------------------------------------------------------*)
IF _bFaultLatch AND bEnable AND bWatchdog AND (NOT tonWd.Q) AND _bCfgOk
   AND (fOutReq = fOutReq) AND (ABS(fOutReq) <= AOF_FIN_MAX) THEN
    _bFaultLatch := FALSE;                     // 清锁存副本（v1.0.1 电平式解除：三成因条件恒可满足）/ clear the latch, level based, always satisfiable
    _uLatch := AOF_ERR_NONE;                   // 清锁存码 / clear the latched code
END_IF

(*------------------------------------------------------------------------------
 * 段 5｜输出映射（名实双出口 R191）：bError/uErrorId 与锁存副本同源
 *      The outlet mapping, the flag and code mirror the latch copy
 *-----------------------------------------------------------------------------*)
IF _bFaultLatch THEN
    bError   := TRUE;                          // 故障标志（R45 配对）/ the fault flag
    uErrorId := _uLatch;                       // 锁存回放 / the latched replay
    IF (_eState = E_DL_AnaOutFsState.eIdle) OR (_eState = E_DL_AnaOutFsState.eNormal) THEN
        _eState := E_DL_AnaOutFsState.eFault;  // 锁存起点迁入故障相（v1.0.1：单次迁入，失保相驻留期不再被回写）/ enter the fault phase at latch onset only
    END_IF
END_IF

(*------------------------------------------------------------------------------
 * 段 6｜状态机（ENUM + CASE，含 ELSE 兜底；eFault 分支显式出现）
 *      The state machine with the else catch all, the fault phase explicit
 *-----------------------------------------------------------------------------*)
IF (NOT bEnable) AND (NOT _bFaultLatch) THEN   // 失能回空闲（v1.0.1：锁存期失保动作优先，不被失能覆盖）/ disable forces idle, the fail action outranks while latched
    _eState := E_DL_AnaOutFsState.eIdle;
END_IF
CASE _eState OF
    E_DL_AnaOutFsState.eIdle:                  // 失能相：输出冻结保持 / the idle phase, output frozen
        IF bEnable AND _bCfgOk AND (NOT _bFaultLatch) THEN
            _eState := E_DL_AnaOutFsState.eNormal;  // 使能迁入正常相 / enter the normal phase on enable
        END_IF
    E_DL_AnaOutFsState.eNormal:                // 正常相：斜坡跟踪请求 / the normal phase, ramp tracking
        IF NOT bEnable THEN
            _eState := E_DL_AnaOutFsState.eIdle;    // 使能撤销回空闲 / back to idle on disable
        ELSIF _bFaultLatch THEN
            _eState := E_DL_AnaOutFsState.eFault;   // 锁存迁入故障相 / enter the fault phase on latch
        ELSE
            IF (fOutReq <> fOutReq) OR (ABS(fOutReq) > AOF_FIN_MAX) THEN
                _fTarget := AOF_OUT_MIN;            // 请求非有限按安全侧下限处理（头注契约）/ a non finite request goes to the safe lower limit
            ELSE
                _bClampReq := FALSE;                // 重置钳位信息位 / reset the clamp flag
                _fTarget := fOutReq;                // 合法请求直取 / take the valid request
                IF _fTarget < AOF_OUT_MIN THEN
                    _fTarget := AOF_OUT_MIN;        // 请求下钳 / clamp the request low
                    _bClampReq := TRUE;             // 记录钳位（信息性）/ mark the clamp
                END_IF
                IF _fTarget > AOF_OUT_MAX THEN
                    _fTarget := AOF_OUT_MAX;        // 请求上钳 / clamp the request high
                    _bClampReq := TRUE;
                END_IF
            END_IF
            _fStep := fRampRatePctS * fCallCycleS;  // 本拍步长 [%]（周期已闸 > 0）/ the per scan step, the cycle gated
            IF fOutAct < _fTarget - 1.0E-9 THEN
                fOutAct := fOutAct + _fStep;        // 向上斜坡 / ramp up
                IF fOutAct > _fTarget THEN fOutAct := _fTarget; END_IF  // 不越过目标 / never past the target
            ELSIF fOutAct > _fTarget + 1.0E-9 THEN
                fOutAct := fOutAct - _fStep;        // 向下斜坡 / ramp down
                IF fOutAct < _fTarget THEN fOutAct := _fTarget; END_IF
            END_IF
        END_IF
    E_DL_AnaOutFsState.eFrozen:                // 失保冻结相：保持当前值（eFreeze 模式落点）/ the fail frozen phase
        IF NOT _bFaultLatch THEN
            _eState := E_DL_AnaOutFsState.eNormal;  // 解除后回正常 / back to normal on release
        ELSIF eFailMode = E_DL_FailMode.eSafeValue THEN
            _eState := E_DL_AnaOutFsState.eSafeHold; // 驻留期切安全值模式：一次完成切换沿 / a mode switch during the dwell lands in one edge
        END_IF
    E_DL_AnaOutFsState.eSafeHold:              // 失保安全值相：斜坡回程到安全值 / the fail safe phase
        IF NOT _bFaultLatch THEN
            _eState := E_DL_AnaOutFsState.eNormal;  // 解除后回正常 / back to normal on release
        ELSIF eFailMode = E_DL_FailMode.eFreeze THEN
            _eState := E_DL_AnaOutFsState.eFrozen;  // 驻留期切冻结模式：一次完成切换沿 / a mode switch during the dwell lands in one edge
        ELSE
            _fStep := fRampRatePctS * fCallCycleS;  // 回程同样限速（斜坡回程限速契约）/ the return path is rate limited too
            IF fOutAct < fSafeValue - 1.0E-9 THEN
                fOutAct := fOutAct + _fStep;
                IF fOutAct > fSafeValue THEN fOutAct := fSafeValue; END_IF
            ELSIF fOutAct > fSafeValue + 1.0E-9 THEN
                fOutAct := fOutAct - _fStep;
                IF fOutAct < fSafeValue THEN fOutAct := fSafeValue; END_IF
            END_IF
        END_IF
    E_DL_AnaOutFsState.eFault:                 // 故障相（显式分支）：按失保模式落冻结/安全值侧
        // eFault 分支动作：本拍按 eFailMode 迁入 eFrozen（保持）或 eSafeHold（回程）；
        // 拍 N 进入故障相 → 本拍完成模式落点 → 拍 N+1 起在对应失保相执行保持/回程
        // the fault phase lands the fail mode in one scan, the hold or ramp runs from the next scan
        IF NOT _bFaultLatch THEN
            _eState := E_DL_AnaOutFsState.eNormal;  // 解除回正常 / back to normal on release
        ELSIF eFailMode = E_DL_FailMode.eFreeze THEN
            _eState := E_DL_AnaOutFsState.eFrozen;  // 冻结模式落点 / land the freeze mode
        ELSE
            _eState := E_DL_AnaOutFsState.eSafeHold; // 安全值模式落点（含非法枚举兜底）/ land the safe mode, also the else style fallback
        END_IF
    ELSE                                        // 非法状态兜底（R 非法态拦截）：落故障相并锁存配置码
        _eState := E_DL_AnaOutFsState.eFault;   // 强制故障相 / force the fault phase
        _bFaultLatch := TRUE;                   // 非法态按锁存处置（R ELSE 兜底不静默）/ an illegal state latches
        _uLatch := AOF_ERR_CFG;
        bError := TRUE;                         // 名实双出口同步 / sync the outlets
        uErrorId := _uLatch;
    END_CASE

(*------------------------------------------------------------------------------
 * 段 7｜输出钳位（双保险切断线）与状态发布 / segment 7, the output clamp and state publish
 *-----------------------------------------------------------------------------*)
IF fOutAct < AOF_OUT_MIN THEN
    fOutAct := AOF_OUT_MIN;                     // 输出下限钳位 / clamp the output low
END_IF
IF fOutAct > AOF_OUT_MAX THEN
    fOutAct := AOF_OUT_MAX;                     // 输出上限钳位 / clamp the output high
END_IF
IF (fOutAct <> fOutAct) THEN                    // 防御：任何路径不得把非有限送出口 / no non finite may reach the outlet
    fOutAct := AOF_OUT_MIN;                     // 落安全下限 / land on the safe lower limit
    _eState := E_DL_AnaOutFsState.eFault;       // 落故障相 / land the fault phase
    _bFaultLatch := TRUE;
    _uLatch := AOF_ERR_REQ;
    bError := TRUE;
    uErrorId := _uLatch;
END_IF
eState := _eState;                              // 状态出口（名实双出口 R191）/ publish the state
END_FUNCTION_BLOCK
